           IF "CNV_HMI".Charge_Commands[#HMI_No] THEN
               CASE #"ID(1)" OF
                       //CNV 1 - SYSTEM 1
                   100101:
                       #"Enable(1)" := "Control_DB".LCnv_Sys[#Sys_No].Cnv_Level[1].Cnv1.Instruction.Enable;
                       #"Mode_Change(1)" := "Control_DB".LCnv_Sys[#Sys_No].Cnv_Level[1].Cnv1.Instruction.Mode_Change;
                       #"Transfer_To_ID(1)" := "Control_DB".LCnv_Sys[#Sys_No].Cnv_Level[1].Cnv1.Instruction.Transfer_To_ID;
                       #"Transfer_From_ID(1)" := "Control_DB".LCnv_Sys[#Sys_No].Cnv_Level[1].Cnv1.Instruction.Transfer_From_ID;
                       #"Pallet_Allignment(1)" := "Control_DB".LCnv_Sys[#Sys_No].Cnv_Level[1].Cnv1.Instruction.Pallet_Allignment;
                   100201:
                       "Enable_HMI(1)" := "Control_DB".LCnv_Sys[#Sys_No].Cnv_Level[2].Cnv1.Instruction.Enable;
                       "Mode_Change_HMI(1)" := "Control_DB".LCnv_Sys[#Sys_No].Cnv_Level[2].Cnv1.Instruction.Mode_Change;
                       "Transfer_To_ID_HMI(1)" := "Control_DB".LCnv_Sys[#Sys_No].Cnv_Level[2].Cnv1.Instruction.Transfer_To_ID;
                       "Transfer_From_ID_HMI(1)" := "Control_DB".LCnv_Sys[#Sys_No].Cnv_Level[2].Cnv1.Instruction.Transfer_From_ID;
                       "Pallet_Allignment_HMI(1)" := "Control_DB".LCnv_Sys[#Sys_No].Cnv_Level[2].Cnv1.Instruction.Pallet_Allignment;
                   100301:
                       "Enable_HMI(1)" := "Control_DB".LCnv_Sys[#Sys_No].Cnv_Level[3].Cnv1.Instruction.Enable;
                       "Mode_Change_HMI(1)" := "Control_DB".LCnv_Sys[#Sys_No].Cnv_Level[3].Cnv1.Instruction.Mode_Change;
                       "Transfer_To_ID_HMI(1)" := "Control_DB".LCnv_Sys[#Sys_No].Cnv_Level[3].Cnv1.Instruction.Transfer_To_ID;
                       "Transfer_From_ID_HMI(1)" := "Control_DB".LCnv_Sys[#Sys_No].Cnv_Level[3].Cnv1.Instruction.Transfer_From_ID;
                       "Pallet_Allignment_HMI(1)" := "Control_DB".LCnv_Sys[#Sys_No].Cnv_Level[3].Cnv1.Instruction.Pallet_Allignment;
                   100401:
                       "Enable_HMI(1)" := "Control_DB".LCnv_Sys[#Sys_No].Cnv_Level[4].Cnv1.Instruction.Enable;
                       "Mode_Change_HMI(1)" := "Control_DB".LCnv_Sys[#Sys_No].Cnv_Level[4].Cnv1.Instruction.Mode_Change;
                       "Transfer_To_ID_HMI(1)" := "Control_DB".LCnv_Sys[#Sys_No].Cnv_Level[4].Cnv1.Instruction.Transfer_To_ID;
                       "Transfer_From_ID_HMI(1)" := "Control_DB".LCnv_Sys[#Sys_No].Cnv_Level[4].Cnv1.Instruction.Transfer_From_ID;
                       "Pallet_Allignment_HMI(1)" := "Control_DB".LCnv_Sys[#Sys_No].Cnv_Level[4].Cnv1.Instruction.Pallet_Allignment;
                   100501:
                       "Enable_HMI(1)" := "Control_DB".LCnv_Sys[#Sys_No].Cnv_Level[5].Cnv1.Instruction.Enable;
                       "Mode_Change_HMI(1)" := "Control_DB".LCnv_Sys[#Sys_No].Cnv_Level[5].Cnv1.Instruction.Mode_Change;
                       "Task_ID_HMI(1)" := "Control_DB".LCnv_Sys[#Sys_No].Cnv_Level[5].Cnv1.Instruction.Task_ID;
                       "Transfer_To_ID_HMI(1)" := "Control_DB".LCnv_Sys[#Sys_No].Cnv_Level[5].Cnv1.Instruction.Transfer_To_ID;
                       "Transfer_From_ID_HMI(1)" := "Control_DB".LCnv_Sys[#Sys_No].Cnv_Level[5].Cnv1.Instruction.Transfer_From_ID;
                       "Pallet_Allignment_HMI(1)" := "Control_DB".LCnv_Sys[#Sys_No].Cnv_Level[5].Cnv1.Instruction.Pallet_Allignment;
                   100601:
                       "Enable_HMI(1)" := "Control_DB".LCnv_Sys[#Sys_No].Cnv_Level[6].Cnv1.Instruction.Enable;
                       "Mode_Change_HMI(1)" := "Control_DB".LCnv_Sys[#Sys_No].Cnv_Level[6].Cnv1.Instruction.Mode_Change;
                       "Task_ID_HMI(1)" := "Control_DB".LCnv_Sys[#Sys_No].Cnv_Level[6].Cnv1.Instruction.Task_ID;
                       "Transfer_To_ID_HMI(1)" := "Control_DB".LCnv_Sys[#Sys_No].Cnv_Level[6].Cnv1.Instruction.Transfer_To_ID;
                       "Transfer_From_ID_HMI(1)" := "Control_DB".LCnv_Sys[#Sys_No].Cnv_Level[6].Cnv1.Instruction.Transfer_From_ID;
                       "Pallet_Allignment_HMI(1)" := "Control_DB".LCnv_Sys[#Sys_No].Cnv_Level[6].Cnv1.Instruction.Pallet_Allignment;
                   100701:
                       "Enable_HMI(1)" := "Control_DB".LCnv_Sys[#Sys_No].Cnv_Level[7].Cnv1.Instruction.Enable;
                       "Mode_Change_HMI(1)" := "Control_DB".LCnv_Sys[#Sys_No].Cnv_Level[7].Cnv1.Instruction.Mode_Change;
                       "Task_ID_HMI(1)" := "Control_DB".LCnv_Sys[#Sys_No].Cnv_Level[7].Cnv1.Instruction.Task_ID;
                       "Transfer_To_ID_HMI(1)" := "Control_DB".LCnv_Sys[#Sys_No].Cnv_Level[7].Cnv1.Instruction.Transfer_To_ID;
                       "Transfer_From_ID_HMI(1)" := "Control_DB".LCnv_Sys[#Sys_No].Cnv_Level[7].Cnv1.Instruction.Transfer_From_ID;
                       "Pallet_Allignment_HMI(1)" := "Control_DB".LCnv_Sys[#Sys_No].Cnv_Level[7].Cnv1.Instruction.Pallet_Allignment;
                   100801:
                       "Enable_HMI(1)" := "Control_DB".LCnv_Sys[#Sys_No].Cnv_Level[8].Cnv1.Instruction.Enable;
                       "Mode_Change_HMI(1)" := "Control_DB".LCnv_Sys[#Sys_No].Cnv_Level[8].Cnv1.Instruction.Mode_Change;
                       "Task_ID_HMI(1)" := "Control_DB".LCnv_Sys[#Sys_No].Cnv_Level[8].Cnv1.Instruction.Task_ID;
                       "Transfer_To_ID_HMI(1)" := "Control_DB".LCnv_Sys[#Sys_No].Cnv_Level[8].Cnv1.Instruction.Transfer_To_ID;
                       "Transfer_From_ID_HMI(1)" := "Control_DB".LCnv_Sys[#Sys_No].Cnv_Level[8].Cnv1.Instruction.Transfer_From_ID;
                       "Pallet_Allignment_HMI(1)" := "Control_DB".LCnv_Sys[#Sys_No].Cnv_Level[8].Cnv1.Instruction.Pallet_Allignment;
                       //CNV 2 - SYSTEM 1
                   110101:
                       "Enable_HMI(1)" := "Control_DB".LCnv_Sys[#Sys_No].Cnv_Level[1].Cnv2.Instruction.Enable;
                       "Mode_Change_HMI(1)" := "Control_DB".LCnv_Sys[#Sys_No].Cnv_Level[1].Cnv2.Instruction.Mode_Change;
                       "Task_ID_HMI(1)" := "Control_DB".LCnv_Sys[#Sys_No].Cnv_Level[1].Cnv2.Instruction.Task_ID;
                       "Transfer_To_ID_HMI(1)" := "Control_DB".LCnv_Sys[#Sys_No].Cnv_Level[1].Cnv2.Instruction.Transfer_To_ID;
                       "Transfer_From_ID_HMI(1)" := "Control_DB".LCnv_Sys[#Sys_No].Cnv_Level[1].Cnv2.Instruction.Transfer_From_ID;
                       "Pallet_Allignment_HMI(1)" := "Control_DB".LCnv_Sys[#Sys_No].Cnv_Level[1].Cnv2.Instruction.Pallet_Allignment;
                   110201:
                       "Enable_HMI(1)" := "Control_DB".LCnv_Sys[#Sys_No].Cnv_Level[2].Cnv2.Instruction.Enable;
                       "Mode_Change_HMI(1)" := "Control_DB".LCnv_Sys[#Sys_No].Cnv_Level[2].Cnv2.Instruction.Mode_Change;
                       "Task_ID_HMI(1)" := "Control_DB".LCnv_Sys[#Sys_No].Cnv_Level[2].Cnv2.Instruction.Task_ID;
                       "Transfer_To_ID_HMI(1)" := "Control_DB".LCnv_Sys[#Sys_No].Cnv_Level[2].Cnv2.Instruction.Transfer_To_ID;
                       "Transfer_From_ID_HMI(1)" := "Control_DB".LCnv_Sys[#Sys_No].Cnv_Level[2].Cnv2.Instruction.Transfer_From_ID;
                       "Pallet_Allignment_HMI(1)" := "Control_DB".LCnv_Sys[#Sys_No].Cnv_Level[2].Cnv2.Instruction.Pallet_Allignment;
                   110301:
                       "Enable_HMI(1)" := "Control_DB".LCnv_Sys[#Sys_No].Cnv_Level[3].Cnv2.Instruction.Enable;
                       "Mode_Change_HMI(1)" := "Control_DB".LCnv_Sys[#Sys_No].Cnv_Level[3].Cnv2.Instruction.Mode_Change;
                       "Task_ID_HMI(1)" := "Control_DB".LCnv_Sys[#Sys_No].Cnv_Level[3].Cnv2.Instruction.Task_ID;
                       "Transfer_To_ID_HMI(1)" := "Control_DB".LCnv_Sys[#Sys_No].Cnv_Level[3].Cnv2.Instruction.Transfer_To_ID;
                       "Transfer_From_ID_HMI(1)" := "Control_DB".LCnv_Sys[#Sys_No].Cnv_Level[3].Cnv2.Instruction.Transfer_From_ID;
                       "Pallet_Allignment_HMI(1)" := "Control_DB".LCnv_Sys[#Sys_No].Cnv_Level[3].Cnv2.Instruction.Pallet_Allignment;
                   110401:
                       "Enable_HMI(1)" := "Control_DB".LCnv_Sys[#Sys_No].Cnv_Level[4].Cnv2.Instruction.Enable;
                       "Mode_Change_HMI(1)" := "Control_DB".LCnv_Sys[#Sys_No].Cnv_Level[4].Cnv2.Instruction.Mode_Change;
                       "Task_ID_HMI(1)" := "Control_DB".LCnv_Sys[#Sys_No].Cnv_Level[4].Cnv2.Instruction.Task_ID;
                       "Transfer_To_ID_HMI(1)" := "Control_DB".LCnv_Sys[#Sys_No].Cnv_Level[4].Cnv2.Instruction.Transfer_To_ID;
                       "Transfer_From_ID_HMI(1)" := "Control_DB".LCnv_Sys[#Sys_No].Cnv_Level[4].Cnv2.Instruction.Transfer_From_ID;
                       "Pallet_Allignment_HMI(1)" := "Control_DB".LCnv_Sys[#Sys_No].Cnv_Level[4].Cnv2.Instruction.Pallet_Allignment;
                   110501:
                       "Enable_HMI(1)" := "Control_DB".LCnv_Sys[#Sys_No].Cnv_Level[5].Cnv2.Instruction.Enable;
                       "Mode_Change_HMI(1)" := "Control_DB".LCnv_Sys[#Sys_No].Cnv_Level[5].Cnv2.Instruction.Mode_Change;
                       "Task_ID_HMI(1)" := "Control_DB".LCnv_Sys[#Sys_No].Cnv_Level[5].Cnv2.Instruction.Task_ID;
                       "Transfer_To_ID_HMI(1)" := "Control_DB".LCnv_Sys[#Sys_No].Cnv_Level[5].Cnv2.Instruction.Transfer_To_ID;
                       "Transfer_From_ID_HMI(1)" := "Control_DB".LCnv_Sys[#Sys_No].Cnv_Level[5].Cnv2.Instruction.Transfer_From_ID;
                       "Pallet_Allignment_HMI(1)" := "Control_DB".LCnv_Sys[#Sys_No].Cnv_Level[5].Cnv2.Instruction.Pallet_Allignment;
                   110601:
                       "Enable_HMI(1)" := "Control_DB".LCnv_Sys[#Sys_No].Cnv_Level[6].Cnv2.Instruction.Enable;
                       "Mode_Change_HMI(1)" := "Control_DB".LCnv_Sys[#Sys_No].Cnv_Level[6].Cnv2.Instruction.Mode_Change;
                       "Task_ID_HMI(1)" := "Control_DB".LCnv_Sys[#Sys_No].Cnv_Level[6].Cnv2.Instruction.Task_ID;
                       "Transfer_To_ID_HMI(1)" := "Control_DB".LCnv_Sys[#Sys_No].Cnv_Level[6].Cnv2.Instruction.Transfer_To_ID;
                       "Transfer_From_ID_HMI(1)" := "Control_DB".LCnv_Sys[#Sys_No].Cnv_Level[6].Cnv2.Instruction.Transfer_From_ID;
                       "Pallet_Allignment_HMI(1)" := "Control_DB".LCnv_Sys[#Sys_No].Cnv_Level[6].Cnv2.Instruction.Pallet_Allignment;
                   110701:
                       "Enable_HMI(1)" := "Control_DB".LCnv_Sys[#Sys_No].Cnv_Level[7].Cnv2.Instruction.Enable;
                       "Mode_Change_HMI(1)" := "Control_DB".LCnv_Sys[#Sys_No].Cnv_Level[7].Cnv2.Instruction.Mode_Change;
                       "Task_ID_HMI(1)" := "Control_DB".LCnv_Sys[#Sys_No].Cnv_Level[7].Cnv2.Instruction.Task_ID;
                       "Transfer_To_ID_HMI(1)" := "Control_DB".LCnv_Sys[#Sys_No].Cnv_Level[7].Cnv2.Instruction.Transfer_To_ID;
                       "Transfer_From_ID_HMI(1)" := "Control_DB".LCnv_Sys[#Sys_No].Cnv_Level[7].Cnv2.Instruction.Transfer_From_ID;
                       "Pallet_Allignment_HMI(1)" := "Control_DB".LCnv_Sys[#Sys_No].Cnv_Level[7].Cnv2.Instruction.Pallet_Allignment;
                   110801:
                       "Enable_HMI(1)" := "Control_DB".LCnv_Sys[#Sys_No].Cnv_Level[8].Cnv2.Instruction.Enable;
                       "Mode_Change_HMI(1)" := "Control_DB".LCnv_Sys[#Sys_No].Cnv_Level[8].Cnv2.Instruction.Mode_Change;
                       "Task_ID_HMI(1)" := "Control_DB".LCnv_Sys[#Sys_No].Cnv_Level[8].Cnv2.Instruction.Task_ID;
                       "Transfer_To_ID_HMI(1)" := "Control_DB".LCnv_Sys[#Sys_No].Cnv_Level[8].Cnv2.Instruction.Transfer_To_ID;
                       "Transfer_From_ID_HMI(1)" := "Control_DB".LCnv_Sys[#Sys_No].Cnv_Level[8].Cnv2.Instruction.Transfer_From_ID;
                       "Pallet_Allignment_HMI(1)" := "Control_DB".LCnv_Sys[#Sys_No].Cnv_Level[8].Cnv2.Instruction.Pallet_Allignment;
                       //CNV 1 - SYSTEM 2
                   100102:
                       "Enable_HMI(1)" := "Control_DB".LCnv_Sys[2].Cnv_Level[1].Cnv1.Instruction.Enable;
                       "Mode_Change_HMI(1)" := "Control_DB".LCnv_Sys[2].Cnv_Level[1].Cnv1.Instruction.Mode_Change;
                       "Task_ID_HMI(1)" := "Control_DB".LCnv_Sys[2].Cnv_Level[1].Cnv1.Instruction.Task_ID;
                       "Transfer_To_ID_HMI(1)" := "Control_DB".LCnv_Sys[2].Cnv_Level[1].Cnv1.Instruction.Transfer_To_ID;
                       "Transfer_From_ID_HMI(1)" := "Control_DB".LCnv_Sys[2].Cnv_Level[1].Cnv1.Instruction.Transfer_From_ID;
                       "Pallet_Allignment_HMI(1)" := "Control_DB".LCnv_Sys[2].Cnv_Level[1].Cnv1.Instruction.Pallet_Allignment;
                   100202:
                       "Enable_HMI(1)" := "Control_DB".LCnv_Sys[2].Cnv_Level[2].Cnv1.Instruction.Enable;
                       "Mode_Change_HMI(1)" := "Control_DB".LCnv_Sys[2].Cnv_Level[2].Cnv1.Instruction.Mode_Change;
                       "Task_ID_HMI(1)" := "Control_DB".LCnv_Sys[2].Cnv_Level[2].Cnv1.Instruction.Task_ID;
                       "Transfer_To_ID_HMI(1)" := "Control_DB".LCnv_Sys[2].Cnv_Level[2].Cnv1.Instruction.Transfer_To_ID;
                       "Transfer_From_ID_HMI(1)" := "Control_DB".LCnv_Sys[2].Cnv_Level[2].Cnv1.Instruction.Transfer_From_ID;
                       "Pallet_Allignment_HMI(1)" := "Control_DB".LCnv_Sys[2].Cnv_Level[2].Cnv1.Instruction.Pallet_Allignment;
                   100302:
                       "Enable_HMI(1)" := "Control_DB".LCnv_Sys[2].Cnv_Level[3].Cnv1.Instruction.Enable;
                       "Mode_Change_HMI(1)" := "Control_DB".LCnv_Sys[2].Cnv_Level[3].Cnv1.Instruction.Mode_Change;
                       "Task_ID_HMI(1)" := "Control_DB".LCnv_Sys[2].Cnv_Level[3].Cnv1.Instruction.Task_ID;
                       "Transfer_To_ID_HMI(1)" := "Control_DB".LCnv_Sys[2].Cnv_Level[3].Cnv1.Instruction.Transfer_To_ID;
                       "Transfer_From_ID_HMI(1)" := "Control_DB".LCnv_Sys[2].Cnv_Level[3].Cnv1.Instruction.Transfer_From_ID;
                       "Pallet_Allignment_HMI(1)" := "Control_DB".LCnv_Sys[2].Cnv_Level[3].Cnv1.Instruction.Pallet_Allignment;
                   100402:
                       "Enable_HMI(1)" := "Control_DB".LCnv_Sys[2].Cnv_Level[4].Cnv1.Instruction.Enable;
                       "Mode_Change_HMI(1)" := "Control_DB".LCnv_Sys[2].Cnv_Level[4].Cnv1.Instruction.Mode_Change;
                       "Task_ID_HMI(1)" := "Control_DB".LCnv_Sys[2].Cnv_Level[4].Cnv1.Instruction.Task_ID;
                       "Transfer_To_ID_HMI(1)" := "Control_DB".LCnv_Sys[2].Cnv_Level[4].Cnv1.Instruction.Transfer_To_ID;
                       "Transfer_From_ID_HMI(1)" := "Control_DB".LCnv_Sys[2].Cnv_Level[4].Cnv1.Instruction.Transfer_From_ID;
                       "Pallet_Allignment_HMI(1)" := "Control_DB".LCnv_Sys[2].Cnv_Level[4].Cnv1.Instruction.Pallet_Allignment;
                   100502:
                       "Enable_HMI(1)" := "Control_DB".LCnv_Sys[2].Cnv_Level[5].Cnv1.Instruction.Enable;
                       "Mode_Change_HMI(1)" := "Control_DB".LCnv_Sys[2].Cnv_Level[5].Cnv1.Instruction.Mode_Change;
                       "Task_ID_HMI(1)" := "Control_DB".LCnv_Sys[2].Cnv_Level[5].Cnv1.Instruction.Task_ID;
                       "Transfer_To_ID_HMI(1)" := "Control_DB".LCnv_Sys[2].Cnv_Level[5].Cnv1.Instruction.Transfer_To_ID;
                       "Transfer_From_ID_HMI(1)" := "Control_DB".LCnv_Sys[2].Cnv_Level[5].Cnv1.Instruction.Transfer_From_ID;
                       "Pallet_Allignment_HMI(1)" := "Control_DB".LCnv_Sys[2].Cnv_Level[5].Cnv1.Instruction.Pallet_Allignment;
                   100602:
                       "Enable_HMI(1)" := "Control_DB".LCnv_Sys[2].Cnv_Level[6].Cnv1.Instruction.Enable;
                       "Mode_Change_HMI(1)" := "Control_DB".LCnv_Sys[2].Cnv_Level[6].Cnv1.Instruction.Mode_Change;
                       "Task_ID_HMI(1)" := "Control_DB".LCnv_Sys[2].Cnv_Level[6].Cnv1.Instruction.Task_ID;
                       "Transfer_To_ID_HMI(1)" := "Control_DB".LCnv_Sys[2].Cnv_Level[6].Cnv1.Instruction.Transfer_To_ID;
                       "Transfer_From_ID_HMI(1)" := "Control_DB".LCnv_Sys[2].Cnv_Level[6].Cnv1.Instruction.Transfer_From_ID;
                       "Pallet_Allignment_HMI(1)" := "Control_DB".LCnv_Sys[2].Cnv_Level[6].Cnv1.Instruction.Pallet_Allignment;
                   100702:
                       "Enable_HMI(1)" := "Control_DB".LCnv_Sys[2].Cnv_Level[7].Cnv1.Instruction.Enable;
                       "Mode_Change_HMI(1)" := "Control_DB".LCnv_Sys[2].Cnv_Level[7].Cnv1.Instruction.Mode_Change;
                       "Task_ID_HMI(1)" := "Control_DB".LCnv_Sys[2].Cnv_Level[7].Cnv1.Instruction.Task_ID;
                       "Transfer_To_ID_HMI(1)" := "Control_DB".LCnv_Sys[2].Cnv_Level[7].Cnv1.Instruction.Transfer_To_ID;
                       "Transfer_From_ID_HMI(1)" := "Control_DB".LCnv_Sys[2].Cnv_Level[7].Cnv1.Instruction.Transfer_From_ID;
                       "Pallet_Allignment_HMI(1)" := "Control_DB".LCnv_Sys[2].Cnv_Level[7].Cnv1.Instruction.Pallet_Allignment;
                   100802:
                       "Enable_HMI(1)" := "Control_DB".LCnv_Sys[2].Cnv_Level[8].Cnv1.Instruction.Enable;
                       "Mode_Change_HMI(1)" := "Control_DB".LCnv_Sys[2].Cnv_Level[8].Cnv1.Instruction.Mode_Change;
                       "Task_ID_HMI(1)" := "Control_DB".LCnv_Sys[2].Cnv_Level[8].Cnv1.Instruction.Task_ID;
                       "Transfer_To_ID_HMI(1)" := "Control_DB".LCnv_Sys[2].Cnv_Level[8].Cnv1.Instruction.Transfer_To_ID;
                       "Transfer_From_ID_HMI(1)" := "Control_DB".LCnv_Sys[2].Cnv_Level[8].Cnv1.Instruction.Transfer_From_ID;
                       "Pallet_Allignment_HMI(1)" := "Control_DB".LCnv_Sys[2].Cnv_Level[8].Cnv1.Instruction.Pallet_Allignment;
                       //CNV 2 - SYSTEM 2
                   110102:
                       "Enable_HMI(1)" := "Control_DB".LCnv_Sys[2].Cnv_Level[1].Cnv2.Instruction.Enable;
                       "Mode_Change_HMI(1)" := "Control_DB".LCnv_Sys[2].Cnv_Level[1].Cnv2.Instruction.Mode_Change;
                       "Task_ID_HMI(1)" := "Control_DB".LCnv_Sys[2].Cnv_Level[1].Cnv2.Instruction.Task_ID;
                       "Transfer_To_ID_HMI(1)" := "Control_DB".LCnv_Sys[2].Cnv_Level[1].Cnv2.Instruction.Transfer_To_ID;
                       "Transfer_From_ID_HMI(1)" := "Control_DB".LCnv_Sys[2].Cnv_Level[1].Cnv2.Instruction.Transfer_From_ID;
                       "Pallet_Allignment_HMI(1)" := "Control_DB".LCnv_Sys[2].Cnv_Level[1].Cnv2.Instruction.Pallet_Allignment;
                   110202:
                       "Enable_HMI(1)" := "Control_DB".LCnv_Sys[2].Cnv_Level[2].Cnv2.Instruction.Enable;
                       "Mode_Change_HMI(1)" := "Control_DB".LCnv_Sys[2].Cnv_Level[2].Cnv2.Instruction.Mode_Change;
                       "Task_ID_HMI(1)" := "Control_DB".LCnv_Sys[2].Cnv_Level[2].Cnv2.Instruction.Task_ID;
                       "Transfer_To_ID_HMI(1)" := "Control_DB".LCnv_Sys[2].Cnv_Level[2].Cnv2.Instruction.Transfer_To_ID;
                       "Transfer_From_ID_HMI(1)" := "Control_DB".LCnv_Sys[2].Cnv_Level[2].Cnv2.Instruction.Transfer_From_ID;
                       "Pallet_Allignment_HMI(1)" := "Control_DB".LCnv_Sys[2].Cnv_Level[2].Cnv2.Instruction.Pallet_Allignment;
                   110302:
                       "Enable_HMI(1)" := "Control_DB".LCnv_Sys[2].Cnv_Level[3].Cnv2.Instruction.Enable;
                       "Mode_Change_HMI(1)" := "Control_DB".LCnv_Sys[2].Cnv_Level[3].Cnv2.Instruction.Mode_Change;
                       "Task_ID_HMI(1)" := "Control_DB".LCnv_Sys[2].Cnv_Level[3].Cnv2.Instruction.Task_ID;
                       "Transfer_To_ID_HMI(1)" := "Control_DB".LCnv_Sys[2].Cnv_Level[3].Cnv2.Instruction.Transfer_To_ID;
                       "Transfer_From_ID_HMI(1)" := "Control_DB".LCnv_Sys[2].Cnv_Level[3].Cnv2.Instruction.Transfer_From_ID;
                       "Pallet_Allignment_HMI(1)" := "Control_DB".LCnv_Sys[2].Cnv_Level[3].Cnv2.Instruction.Pallet_Allignment;
                   110402:
                       "Enable_HMI(1)" := "Control_DB".LCnv_Sys[2].Cnv_Level[4].Cnv2.Instruction.Enable;
                       "Mode_Change_HMI(1)" := "Control_DB".LCnv_Sys[2].Cnv_Level[4].Cnv2.Instruction.Mode_Change;
                       "Task_ID_HMI(1)" := "Control_DB".LCnv_Sys[2].Cnv_Level[4].Cnv2.Instruction.Task_ID;
                       "Transfer_To_ID_HMI(1)" := "Control_DB".LCnv_Sys[2].Cnv_Level[4].Cnv2.Instruction.Transfer_To_ID;
                       "Transfer_From_ID_HMI(1)" := "Control_DB".LCnv_Sys[2].Cnv_Level[4].Cnv2.Instruction.Transfer_From_ID;
                       "Pallet_Allignment_HMI(1)" := "Control_DB".LCnv_Sys[2].Cnv_Level[4].Cnv2.Instruction.Pallet_Allignment;
                   110502:
                       "Enable_HMI(1)" := "Control_DB".LCnv_Sys[2].Cnv_Level[5].Cnv2.Instruction.Enable;
                       "Mode_Change_HMI(1)" := "Control_DB".LCnv_Sys[2].Cnv_Level[5].Cnv2.Instruction.Mode_Change;
                       "Task_ID_HMI(1)" := "Control_DB".LCnv_Sys[2].Cnv_Level[5].Cnv2.Instruction.Task_ID;
                       "Transfer_To_ID_HMI(1)" := "Control_DB".LCnv_Sys[2].Cnv_Level[5].Cnv2.Instruction.Transfer_To_ID;
                       "Transfer_From_ID_HMI(1)" := "Control_DB".LCnv_Sys[2].Cnv_Level[5].Cnv2.Instruction.Transfer_From_ID;
                       "Pallet_Allignment_HMI(1)" := "Control_DB".LCnv_Sys[2].Cnv_Level[5].Cnv2.Instruction.Pallet_Allignment;
                   110602:
                       "Enable_HMI(1)" := "Control_DB".LCnv_Sys[2].Cnv_Level[6].Cnv2.Instruction.Enable;
                       "Mode_Change_HMI(1)" := "Control_DB".LCnv_Sys[2].Cnv_Level[6].Cnv2.Instruction.Mode_Change;
                       "Task_ID_HMI(1)" := "Control_DB".LCnv_Sys[2].Cnv_Level[6].Cnv2.Instruction.Task_ID;
                       "Transfer_To_ID_HMI(1)" := "Control_DB".LCnv_Sys[2].Cnv_Level[6].Cnv2.Instruction.Transfer_To_ID;
                       "Transfer_From_ID_HMI(1)" := "Control_DB".LCnv_Sys[2].Cnv_Level[6].Cnv2.Instruction.Transfer_From_ID;
                       "Pallet_Allignment_HMI(1)" := "Control_DB".LCnv_Sys[2].Cnv_Level[6].Cnv2.Instruction.Pallet_Allignment;
                   110702:
                       "Enable_HMI(1)" := "Control_DB".LCnv_Sys[2].Cnv_Level[7].Cnv2.Instruction.Enable;
                       "Mode_Change_HMI(1)" := "Control_DB".LCnv_Sys[2].Cnv_Level[7].Cnv2.Instruction.Mode_Change;
                       "Task_ID_HMI(1)" := "Control_DB".LCnv_Sys[2].Cnv_Level[7].Cnv2.Instruction.Task_ID;
                       "Transfer_To_ID_HMI(1)" := "Control_DB".LCnv_Sys[2].Cnv_Level[7].Cnv2.Instruction.Transfer_To_ID;
                       "Transfer_From_ID_HMI(1)" := "Control_DB".LCnv_Sys[2].Cnv_Level[7].Cnv2.Instruction.Transfer_From_ID;
                       "Pallet_Allignment_HMI(1)" := "Control_DB".LCnv_Sys[2].Cnv_Level[7].Cnv2.Instruction.Pallet_Allignment;
                   110802:
                       "Enable_HMI(1)" := "Control_DB".LCnv_Sys[2].Cnv_Level[8].Cnv2.Instruction.Enable;
                       "Mode_Change_HMI(1)" := "Control_DB".LCnv_Sys[2].Cnv_Level[8].Cnv2.Instruction.Mode_Change;
                       "Task_ID_HMI(1)" := "Control_DB".LCnv_Sys[2].Cnv_Level[8].Cnv2.Instruction.Task_ID;
                       "Transfer_To_ID_HMI(1)" := "Control_DB".LCnv_Sys[2].Cnv_Level[8].Cnv2.Instruction.Transfer_To_ID;
                       "Transfer_From_ID_HMI(1)" := "Control_DB".LCnv_Sys[2].Cnv_Level[8].Cnv2.Instruction.Transfer_From_ID;
                       "Pallet_Allignment_HMI(1)" := "Control_DB".LCnv_Sys[2].Cnv_Level[8].Cnv2.Instruction.Pallet_Allignment;
                       //CNV 1 - SYSTEM 3
                   100103:
                       "Enable_HMI(1)" := "Control_DB".LCnv_Sys[3].Cnv_Level[1].Cnv1.Instruction.Enable;
                       "Mode_Change_HMI(1)" := "Control_DB".LCnv_Sys[3].Cnv_Level[1].Cnv1.Instruction.Mode_Change;
                       "Task_ID_HMI(1)" := "Control_DB".LCnv_Sys[3].Cnv_Level[1].Cnv1.Instruction.Task_ID;
                       "Transfer_To_ID_HMI(1)" := "Control_DB".LCnv_Sys[3].Cnv_Level[1].Cnv1.Instruction.Transfer_To_ID;
                       "Transfer_From_ID_HMI(1)" := "Control_DB".LCnv_Sys[3].Cnv_Level[1].Cnv1.Instruction.Transfer_From_ID;
                       "Pallet_Allignment_HMI(1)" := "Control_DB".LCnv_Sys[3].Cnv_Level[1].Cnv1.Instruction.Pallet_Allignment;
                   100203:
                       "Enable_HMI(1)" := "Control_DB".LCnv_Sys[3].Cnv_Level[2].Cnv1.Instruction.Enable;
                       "Mode_Change_HMI(1)" := "Control_DB".LCnv_Sys[3].Cnv_Level[2].Cnv1.Instruction.Mode_Change;
                       "Task_ID_HMI(1)" := "Control_DB".LCnv_Sys[3].Cnv_Level[2].Cnv1.Instruction.Task_ID;
                       "Transfer_To_ID_HMI(1)" := "Control_DB".LCnv_Sys[3].Cnv_Level[2].Cnv1.Instruction.Transfer_To_ID;
                       "Transfer_From_ID_HMI(1)" := "Control_DB".LCnv_Sys[3].Cnv_Level[2].Cnv1.Instruction.Transfer_From_ID;
                       "Pallet_Allignment_HMI(1)" := "Control_DB".LCnv_Sys[3].Cnv_Level[2].Cnv1.Instruction.Pallet_Allignment;
                   100303:
                       "Enable_HMI(1)" := "Control_DB".LCnv_Sys[3].Cnv_Level[3].Cnv1.Instruction.Enable;
                       "Mode_Change_HMI(1)" := "Control_DB".LCnv_Sys[3].Cnv_Level[3].Cnv1.Instruction.Mode_Change;
                       "Task_ID_HMI(1)" := "Control_DB".LCnv_Sys[3].Cnv_Level[3].Cnv1.Instruction.Task_ID;
                       "Transfer_To_ID_HMI(1)" := "Control_DB".LCnv_Sys[3].Cnv_Level[3].Cnv1.Instruction.Transfer_To_ID;
                       "Transfer_From_ID_HMI(1)" := "Control_DB".LCnv_Sys[3].Cnv_Level[3].Cnv1.Instruction.Transfer_From_ID;
                       "Pallet_Allignment_HMI(1)" := "Control_DB".LCnv_Sys[3].Cnv_Level[3].Cnv1.Instruction.Pallet_Allignment;
                   100403:
                       "Enable_HMI(1)" := "Control_DB".LCnv_Sys[3].Cnv_Level[4].Cnv1.Instruction.Enable;
                       "Mode_Change_HMI(1)" := "Control_DB".LCnv_Sys[3].Cnv_Level[4].Cnv1.Instruction.Mode_Change;
                       "Task_ID_HMI(1)" := "Control_DB".LCnv_Sys[3].Cnv_Level[4].Cnv1.Instruction.Task_ID;
                       "Transfer_To_ID_HMI(1)" := "Control_DB".LCnv_Sys[3].Cnv_Level[4].Cnv1.Instruction.Transfer_To_ID;
                       "Transfer_From_ID_HMI(1)" := "Control_DB".LCnv_Sys[3].Cnv_Level[4].Cnv1.Instruction.Transfer_From_ID;
                       "Pallet_Allignment_HMI(1)" := "Control_DB".LCnv_Sys[3].Cnv_Level[4].Cnv1.Instruction.Pallet_Allignment;
                   100503:
                       "Enable_HMI(1)" := "Control_DB".LCnv_Sys[3].Cnv_Level[5].Cnv1.Instruction.Enable;
                       "Mode_Change_HMI(1)" := "Control_DB".LCnv_Sys[3].Cnv_Level[5].Cnv1.Instruction.Mode_Change;
                       "Task_ID_HMI(1)" := "Control_DB".LCnv_Sys[3].Cnv_Level[5].Cnv1.Instruction.Task_ID;
                       "Transfer_To_ID_HMI(1)" := "Control_DB".LCnv_Sys[3].Cnv_Level[5].Cnv1.Instruction.Transfer_To_ID;
                       "Transfer_From_ID_HMI(1)" := "Control_DB".LCnv_Sys[3].Cnv_Level[5].Cnv1.Instruction.Transfer_From_ID;
                       "Pallet_Allignment_HMI(1)" := "Control_DB".LCnv_Sys[3].Cnv_Level[5].Cnv1.Instruction.Pallet_Allignment;
                   100603:
                       "Enable_HMI(1)" := "Control_DB".LCnv_Sys[3].Cnv_Level[6].Cnv1.Instruction.Enable;
                       "Mode_Change_HMI(1)" := "Control_DB".LCnv_Sys[3].Cnv_Level[6].Cnv1.Instruction.Mode_Change;
                       "Task_ID_HMI(1)" := "Control_DB".LCnv_Sys[3].Cnv_Level[6].Cnv1.Instruction.Task_ID;
                       "Transfer_To_ID_HMI(1)" := "Control_DB".LCnv_Sys[3].Cnv_Level[6].Cnv1.Instruction.Transfer_To_ID;
                       "Transfer_From_ID_HMI(1)" := "Control_DB".LCnv_Sys[3].Cnv_Level[6].Cnv1.Instruction.Transfer_From_ID;
                       "Pallet_Allignment_HMI(1)" := "Control_DB".LCnv_Sys[3].Cnv_Level[6].Cnv1.Instruction.Pallet_Allignment;
                   100703:
                       "Enable_HMI(1)" := "Control_DB".LCnv_Sys[3].Cnv_Level[7].Cnv1.Instruction.Enable;
                       "Mode_Change_HMI(1)" := "Control_DB".LCnv_Sys[3].Cnv_Level[7].Cnv1.Instruction.Mode_Change;
                       "Task_ID_HMI(1)" := "Control_DB".LCnv_Sys[3].Cnv_Level[7].Cnv1.Instruction.Task_ID;
                       "Transfer_To_ID_HMI(1)" := "Control_DB".LCnv_Sys[3].Cnv_Level[7].Cnv1.Instruction.Transfer_To_ID;
                       "Transfer_From_ID_HMI(1)" := "Control_DB".LCnv_Sys[3].Cnv_Level[7].Cnv1.Instruction.Transfer_From_ID;
                       "Pallet_Allignment_HMI(1)" := "Control_DB".LCnv_Sys[3].Cnv_Level[7].Cnv1.Instruction.Pallet_Allignment;
                   100803:
                       "Enable_HMI(1)" := "Control_DB".LCnv_Sys[3].Cnv_Level[8].Cnv1.Instruction.Enable;
                       "Mode_Change_HMI(1)" := "Control_DB".LCnv_Sys[3].Cnv_Level[8].Cnv1.Instruction.Mode_Change;
                       "Task_ID_HMI(1)" := "Control_DB".LCnv_Sys[3].Cnv_Level[8].Cnv1.Instruction.Task_ID;
                       "Transfer_To_ID_HMI(1)" := "Control_DB".LCnv_Sys[3].Cnv_Level[8].Cnv1.Instruction.Transfer_To_ID;
                       "Transfer_From_ID_HMI(1)" := "Control_DB".LCnv_Sys[3].Cnv_Level[8].Cnv1.Instruction.Transfer_From_ID;
                       "Pallet_Allignment_HMI(1)" := "Control_DB".LCnv_Sys[3].Cnv_Level[8].Cnv1.Instruction.Pallet_Allignment;
                       //CNV 2 - SYSTEM 3
                   110103:
                       "Enable_HMI(1)" := "Control_DB".LCnv_Sys[3].Cnv_Level[1].Cnv2.Instruction.Enable;
                       "Mode_Change_HMI(1)" := "Control_DB".LCnv_Sys[3].Cnv_Level[1].Cnv2.Instruction.Mode_Change;
                       "Task_ID_HMI(1)" := "Control_DB".LCnv_Sys[3].Cnv_Level[1].Cnv2.Instruction.Task_ID;
                       "Transfer_To_ID_HMI(1)" := "Control_DB".LCnv_Sys[3].Cnv_Level[1].Cnv2.Instruction.Transfer_To_ID;
                       "Transfer_From_ID_HMI(1)" := "Control_DB".LCnv_Sys[3].Cnv_Level[1].Cnv2.Instruction.Transfer_From_ID;
                       "Pallet_Allignment_HMI(1)" := "Control_DB".LCnv_Sys[3].Cnv_Level[1].Cnv2.Instruction.Pallet_Allignment;
                   110203:
                       "Enable_HMI(1)" := "Control_DB".LCnv_Sys[3].Cnv_Level[2].Cnv2.Instruction.Enable;
                       "Mode_Change_HMI(1)" := "Control_DB".LCnv_Sys[3].Cnv_Level[2].Cnv2.Instruction.Mode_Change;
                       "Task_ID_HMI(1)" := "Control_DB".LCnv_Sys[3].Cnv_Level[2].Cnv2.Instruction.Task_ID;
                       "Transfer_To_ID_HMI(1)" := "Control_DB".LCnv_Sys[3].Cnv_Level[2].Cnv2.Instruction.Transfer_To_ID;
                       "Transfer_From_ID_HMI(1)" := "Control_DB".LCnv_Sys[3].Cnv_Level[2].Cnv2.Instruction.Transfer_From_ID;
                       "Pallet_Allignment_HMI(1)" := "Control_DB".LCnv_Sys[3].Cnv_Level[2].Cnv2.Instruction.Pallet_Allignment;
                   110303:
                       "Enable_HMI(1)" := "Control_DB".LCnv_Sys[3].Cnv_Level[3].Cnv2.Instruction.Enable;
                       "Mode_Change_HMI(1)" := "Control_DB".LCnv_Sys[3].Cnv_Level[3].Cnv2.Instruction.Mode_Change;
                       "Task_ID_HMI(1)" := "Control_DB".LCnv_Sys[3].Cnv_Level[3].Cnv2.Instruction.Task_ID;
                       "Transfer_To_ID_HMI(1)" := "Control_DB".LCnv_Sys[3].Cnv_Level[3].Cnv2.Instruction.Transfer_To_ID;
                       "Transfer_From_ID_HMI(1)" := "Control_DB".LCnv_Sys[3].Cnv_Level[3].Cnv2.Instruction.Transfer_From_ID;
                       "Pallet_Allignment_HMI(1)" := "Control_DB".LCnv_Sys[3].Cnv_Level[3].Cnv2.Instruction.Pallet_Allignment;
                   110403:
                       "Enable_HMI(1)" := "Control_DB".LCnv_Sys[3].Cnv_Level[4].Cnv2.Instruction.Enable;
                       "Mode_Change_HMI(1)" := "Control_DB".LCnv_Sys[3].Cnv_Level[4].Cnv2.Instruction.Mode_Change;
                       "Task_ID_HMI(1)" := "Control_DB".LCnv_Sys[3].Cnv_Level[4].Cnv2.Instruction.Task_ID;
                       "Transfer_To_ID_HMI(1)" := "Control_DB".LCnv_Sys[3].Cnv_Level[4].Cnv2.Instruction.Transfer_To_ID;
                       "Transfer_From_ID_HMI(1)" := "Control_DB".LCnv_Sys[3].Cnv_Level[4].Cnv2.Instruction.Transfer_From_ID;
                       "Pallet_Allignment_HMI(1)" := "Control_DB".LCnv_Sys[3].Cnv_Level[4].Cnv2.Instruction.Pallet_Allignment;
                   110503:
                       "Enable_HMI(1)" := "Control_DB".LCnv_Sys[3].Cnv_Level[5].Cnv2.Instruction.Enable;
                       "Mode_Change_HMI(1)" := "Control_DB".LCnv_Sys[3].Cnv_Level[5].Cnv2.Instruction.Mode_Change;
                       "Task_ID_HMI(1)" := "Control_DB".LCnv_Sys[3].Cnv_Level[5].Cnv2.Instruction.Task_ID;
                       "Transfer_To_ID_HMI(1)" := "Control_DB".LCnv_Sys[3].Cnv_Level[5].Cnv2.Instruction.Transfer_To_ID;
                       "Transfer_From_ID_HMI(1)" := "Control_DB".LCnv_Sys[3].Cnv_Level[5].Cnv2.Instruction.Transfer_From_ID;
                       "Pallet_Allignment_HMI(1)" := "Control_DB".LCnv_Sys[3].Cnv_Level[5].Cnv2.Instruction.Pallet_Allignment;
                   110603:
                       "Enable_HMI(1)" := "Control_DB".LCnv_Sys[3].Cnv_Level[6].Cnv2.Instruction.Enable;
                       "Mode_Change_HMI(1)" := "Control_DB".LCnv_Sys[3].Cnv_Level[6].Cnv2.Instruction.Mode_Change;
                       "Task_ID_HMI(1)" := "Control_DB".LCnv_Sys[3].Cnv_Level[6].Cnv2.Instruction.Task_ID;
                       "Transfer_To_ID_HMI(1)" := "Control_DB".LCnv_Sys[3].Cnv_Level[6].Cnv2.Instruction.Transfer_To_ID;
                       "Transfer_From_ID_HMI(1)" := "Control_DB".LCnv_Sys[3].Cnv_Level[6].Cnv2.Instruction.Transfer_From_ID;
                       "Pallet_Allignment_HMI(1)" := "Control_DB".LCnv_Sys[3].Cnv_Level[6].Cnv2.Instruction.Pallet_Allignment;
                   110703:
                       "Enable_HMI(1)" := "Control_DB".LCnv_Sys[3].Cnv_Level[7].Cnv2.Instruction.Enable;
                       "Mode_Change_HMI(1)" := "Control_DB".LCnv_Sys[3].Cnv_Level[7].Cnv2.Instruction.Mode_Change;
                       "Task_ID_HMI(1)" := "Control_DB".LCnv_Sys[3].Cnv_Level[7].Cnv2.Instruction.Task_ID;
                       "Transfer_To_ID_HMI(1)" := "Control_DB".LCnv_Sys[3].Cnv_Level[7].Cnv2.Instruction.Transfer_To_ID;
                       "Transfer_From_ID_HMI(1)" := "Control_DB".LCnv_Sys[3].Cnv_Level[7].Cnv2.Instruction.Transfer_From_ID;
                       "Pallet_Allignment_HMI(1)" := "Control_DB".LCnv_Sys[3].Cnv_Level[7].Cnv2.Instruction.Pallet_Allignment;
                   110803:
                       "Enable_HMI(1)" := "Control_DB".LCnv_Sys[3].Cnv_Level[8].Cnv2.Instruction.Enable;
                       "Mode_Change_HMI(1)" := "Control_DB".LCnv_Sys[3].Cnv_Level[8].Cnv2.Instruction.Mode_Change;
                       "Task_ID_HMI(1)" := "Control_DB".LCnv_Sys[3].Cnv_Level[8].Cnv2.Instruction.Task_ID;
                       "Transfer_To_ID_HMI(1)" := "Control_DB".LCnv_Sys[3].Cnv_Level[8].Cnv2.Instruction.Transfer_To_ID;
                       "Transfer_From_ID_HMI(1)" := "Control_DB".LCnv_Sys[3].Cnv_Level[8].Cnv2.Instruction.Transfer_From_ID;
                       "Pallet_Allignment_HMI(1)" := "Control_DB".LCnv_Sys[3].Cnv_Level[8].Cnv2.Instruction.Pallet_Allignment;
                       //CNV 2 - SYSTEM 4
                   110104:
                       "Enable_HMI(1)" := "Control_DB".LCnv_Sys[4].Cnv_Level[1].Cnv2.Instruction.Enable;
                       "Mode_Change_HMI(1)" := "Control_DB".LCnv_Sys[4].Cnv_Level[1].Cnv2.Instruction.Mode_Change;
                       "Task_ID_HMI(1)" := "Control_DB".LCnv_Sys[4].Cnv_Level[1].Cnv2.Instruction.Task_ID;
                       "Transfer_To_ID_HMI(1)" := "Control_DB".LCnv_Sys[4].Cnv_Level[1].Cnv2.Instruction.Transfer_To_ID;
                       "Transfer_From_ID_HMI(1)" := "Control_DB".LCnv_Sys[4].Cnv_Level[1].Cnv2.Instruction.Transfer_From_ID;
                       "Pallet_Allignment_HMI(1)" := "Control_DB".LCnv_Sys[4].Cnv_Level[1].Cnv2.Instruction.Pallet_Allignment;
                   110204:
                       "Enable_HMI(1)" := "Control_DB".LCnv_Sys[4].Cnv_Level[2].Cnv2.Instruction.Enable;
                       "Mode_Change_HMI(1)" := "Control_DB".LCnv_Sys[4].Cnv_Level[2].Cnv2.Instruction.Mode_Change;
                       "Task_ID_HMI(1)" := "Control_DB".LCnv_Sys[4].Cnv_Level[2].Cnv2.Instruction.Task_ID;
                       "Transfer_To_ID_HMI(1)" := "Control_DB".LCnv_Sys[4].Cnv_Level[2].Cnv2.Instruction.Transfer_To_ID;
                       "Transfer_From_ID_HMI(1)" := "Control_DB".LCnv_Sys[4].Cnv_Level[2].Cnv2.Instruction.Transfer_From_ID;
                       "Pallet_Allignment_HMI(1)" := "Control_DB".LCnv_Sys[4].Cnv_Level[2].Cnv2.Instruction.Pallet_Allignment;
                   110304:
                       "Enable_HMI(1)" := "Control_DB".LCnv_Sys[4].Cnv_Level[3].Cnv2.Instruction.Enable;
                       "Mode_Change_HMI(1)" := "Control_DB".LCnv_Sys[4].Cnv_Level[3].Cnv2.Instruction.Mode_Change;
                       "Task_ID_HMI(1)" := "Control_DB".LCnv_Sys[4].Cnv_Level[3].Cnv2.Instruction.Task_ID;
                       "Transfer_To_ID_HMI(1)" := "Control_DB".LCnv_Sys[4].Cnv_Level[3].Cnv2.Instruction.Transfer_To_ID;
                       "Transfer_From_ID_HMI(1)" := "Control_DB".LCnv_Sys[4].Cnv_Level[3].Cnv2.Instruction.Transfer_From_ID;
                       "Pallet_Allignment_HMI(1)" := "Control_DB".LCnv_Sys[4].Cnv_Level[3].Cnv2.Instruction.Pallet_Allignment;
                   110404:
                       "Enable_HMI(1)" := "Control_DB".LCnv_Sys[4].Cnv_Level[4].Cnv2.Instruction.Enable;
                       "Mode_Change_HMI(1)" := "Control_DB".LCnv_Sys[4].Cnv_Level[4].Cnv2.Instruction.Mode_Change;
                       "Task_ID_HMI(1)" := "Control_DB".LCnv_Sys[4].Cnv_Level[4].Cnv2.Instruction.Task_ID;
                       "Transfer_To_ID_HMI(1)" := "Control_DB".LCnv_Sys[4].Cnv_Level[4].Cnv2.Instruction.Transfer_To_ID;
                       "Transfer_From_ID_HMI(1)" := "Control_DB".LCnv_Sys[4].Cnv_Level[4].Cnv2.Instruction.Transfer_From_ID;
                       "Pallet_Allignment_HMI(1)" := "Control_DB".LCnv_Sys[4].Cnv_Level[4].Cnv2.Instruction.Pallet_Allignment;
                   110504:
                       "Enable_HMI(1)" := "Control_DB".LCnv_Sys[4].Cnv_Level[5].Cnv2.Instruction.Enable;
                       "Mode_Change_HMI(1)" := "Control_DB".LCnv_Sys[4].Cnv_Level[5].Cnv2.Instruction.Mode_Change;
                       "Task_ID_HMI(1)" := "Control_DB".LCnv_Sys[4].Cnv_Level[5].Cnv2.Instruction.Task_ID;
                       "Transfer_To_ID_HMI(1)" := "Control_DB".LCnv_Sys[4].Cnv_Level[5].Cnv2.Instruction.Transfer_To_ID;
                       "Transfer_From_ID_HMI(1)" := "Control_DB".LCnv_Sys[4].Cnv_Level[5].Cnv2.Instruction.Transfer_From_ID;
                       "Pallet_Allignment_HMI(1)" := "Control_DB".LCnv_Sys[4].Cnv_Level[5].Cnv2.Instruction.Pallet_Allignment;
                   110604:
                       "Enable_HMI(1)" := "Control_DB".LCnv_Sys[4].Cnv_Level[6].Cnv2.Instruction.Enable;
                       "Mode_Change_HMI(1)" := "Control_DB".LCnv_Sys[4].Cnv_Level[6].Cnv2.Instruction.Mode_Change;
                       "Task_ID_HMI(1)" := "Control_DB".LCnv_Sys[4].Cnv_Level[6].Cnv2.Instruction.Task_ID;
                       "Transfer_To_ID_HMI(1)" := "Control_DB".LCnv_Sys[4].Cnv_Level[6].Cnv2.Instruction.Transfer_To_ID;
                       "Transfer_From_ID_HMI(1)" := "Control_DB".LCnv_Sys[4].Cnv_Level[6].Cnv2.Instruction.Transfer_From_ID;
                       "Pallet_Allignment_HMI(1)" := "Control_DB".LCnv_Sys[4].Cnv_Level[6].Cnv2.Instruction.Pallet_Allignment;
                   110704:
                       "Enable_HMI(1)" := "Control_DB".LCnv_Sys[4].Cnv_Level[7].Cnv2.Instruction.Enable;
                       "Mode_Change_HMI(1)" := "Control_DB".LCnv_Sys[4].Cnv_Level[7].Cnv2.Instruction.Mode_Change;
                       "Task_ID_HMI(1)" := "Control_DB".LCnv_Sys[4].Cnv_Level[7].Cnv2.Instruction.Task_ID;
                       "Transfer_To_ID_HMI(1)" := "Control_DB".LCnv_Sys[4].Cnv_Level[7].Cnv2.Instruction.Transfer_To_ID;
                       "Transfer_From_ID_HMI(1)" := "Control_DB".LCnv_Sys[4].Cnv_Level[7].Cnv2.Instruction.Transfer_From_ID;
                       "Pallet_Allignment_HMI(1)" := "Control_DB".LCnv_Sys[4].Cnv_Level[7].Cnv2.Instruction.Pallet_Allignment;
                   110804:
                       "Enable_HMI(1)" := "Control_DB".LCnv_Sys[4].Cnv_Level[8].Cnv2.Instruction.Enable;
                       "Mode_Change_HMI(1)" := "Control_DB".LCnv_Sys[4].Cnv_Level[8].Cnv2.Instruction.Mode_Change;
                       "Task_ID_HMI(1)" := "Control_DB".LCnv_Sys[4].Cnv_Level[8].Cnv2.Instruction.Task_ID;
                       "Transfer_To_ID_HMI(1)" := "Control_DB".LCnv_Sys[4].Cnv_Level[8].Cnv2.Instruction.Transfer_To_ID;
                       "Transfer_From_ID_HMI(1)" := "Control_DB".LCnv_Sys[4].Cnv_Level[8].Cnv2.Instruction.Transfer_From_ID;
                       "Pallet_Allignment_HMI(1)" := "Control_DB".LCnv_Sys[4].Cnv_Level[8].Cnv2.Instruction.Pallet_Allignment;
                       //CNV 2 - SYSTEM 5
                   110105:
                       "Enable_HMI(1)" := "Control_DB".LCnv_Sys[5].Cnv_Level[1].Cnv2.Instruction.Enable;
                       "Mode_Change_HMI(1)" := "Control_DB".LCnv_Sys[5].Cnv_Level[1].Cnv2.Instruction.Mode_Change;
                       "Task_ID_HMI(1)" := "Control_DB".LCnv_Sys[5].Cnv_Level[1].Cnv2.Instruction.Task_ID;
                       "Transfer_To_ID_HMI(1)" := "Control_DB".LCnv_Sys[5].Cnv_Level[1].Cnv2.Instruction.Transfer_To_ID;
                       "Transfer_From_ID_HMI(1)" := "Control_DB".LCnv_Sys[5].Cnv_Level[1].Cnv2.Instruction.Transfer_From_ID;
                       "Pallet_Allignment_HMI(1)" := "Control_DB".LCnv_Sys[5].Cnv_Level[1].Cnv2.Instruction.Pallet_Allignment;
                   110205:
                       "Enable_HMI(1)" := "Control_DB".LCnv_Sys[5].Cnv_Level[2].Cnv2.Instruction.Enable;
                       "Mode_Change_HMI(1)" := "Control_DB".LCnv_Sys[5].Cnv_Level[2].Cnv2.Instruction.Mode_Change;
                       "Task_ID_HMI(1)" := "Control_DB".LCnv_Sys[5].Cnv_Level[2].Cnv2.Instruction.Task_ID;
                       "Transfer_To_ID_HMI(1)" := "Control_DB".LCnv_Sys[5].Cnv_Level[2].Cnv2.Instruction.Transfer_To_ID;
                       "Transfer_From_ID_HMI(1)" := "Control_DB".LCnv_Sys[5].Cnv_Level[2].Cnv2.Instruction.Transfer_From_ID;
                       "Pallet_Allignment_HMI(1)" := "Control_DB".LCnv_Sys[5].Cnv_Level[2].Cnv2.Instruction.Pallet_Allignment;
                   110305:
                       "Enable_HMI(1)" := "Control_DB".LCnv_Sys[5].Cnv_Level[3].Cnv2.Instruction.Enable;
                       "Mode_Change_HMI(1)" := "Control_DB".LCnv_Sys[5].Cnv_Level[3].Cnv2.Instruction.Mode_Change;
                       "Task_ID_HMI(1)" := "Control_DB".LCnv_Sys[5].Cnv_Level[3].Cnv2.Instruction.Task_ID;
                       "Transfer_To_ID_HMI(1)" := "Control_DB".LCnv_Sys[5].Cnv_Level[3].Cnv2.Instruction.Transfer_To_ID;
                       "Transfer_From_ID_HMI(1)" := "Control_DB".LCnv_Sys[5].Cnv_Level[3].Cnv2.Instruction.Transfer_From_ID;
                       "Pallet_Allignment_HMI(1)" := "Control_DB".LCnv_Sys[5].Cnv_Level[3].Cnv2.Instruction.Pallet_Allignment;
                   110405:
                       "Enable_HMI(1)" := "Control_DB".LCnv_Sys[5].Cnv_Level[4].Cnv2.Instruction.Enable;
                       "Mode_Change_HMI(1)" := "Control_DB".LCnv_Sys[5].Cnv_Level[4].Cnv2.Instruction.Mode_Change;
                       "Task_ID_HMI(1)" := "Control_DB".LCnv_Sys[5].Cnv_Level[4].Cnv2.Instruction.Task_ID;
                       "Transfer_To_ID_HMI(1)" := "Control_DB".LCnv_Sys[5].Cnv_Level[4].Cnv2.Instruction.Transfer_To_ID;
                       "Transfer_From_ID_HMI(1)" := "Control_DB".LCnv_Sys[5].Cnv_Level[4].Cnv2.Instruction.Transfer_From_ID;
                       "Pallet_Allignment_HMI(1)" := "Control_DB".LCnv_Sys[5].Cnv_Level[4].Cnv2.Instruction.Pallet_Allignment;
                   110505:
                       "Enable_HMI(1)" := "Control_DB".LCnv_Sys[5].Cnv_Level[5].Cnv2.Instruction.Enable;
                       "Mode_Change_HMI(1)" := "Control_DB".LCnv_Sys[5].Cnv_Level[5].Cnv2.Instruction.Mode_Change;
                       "Task_ID_HMI(1)" := "Control_DB".LCnv_Sys[5].Cnv_Level[5].Cnv2.Instruction.Task_ID;
                       "Transfer_To_ID_HMI(1)" := "Control_DB".LCnv_Sys[5].Cnv_Level[5].Cnv2.Instruction.Transfer_To_ID;
                       "Transfer_From_ID_HMI(1)" := "Control_DB".LCnv_Sys[5].Cnv_Level[5].Cnv2.Instruction.Transfer_From_ID;
                       "Pallet_Allignment_HMI(1)" := "Control_DB".LCnv_Sys[5].Cnv_Level[5].Cnv2.Instruction.Pallet_Allignment;
                   110605:
                       "Enable_HMI(1)" := "Control_DB".LCnv_Sys[5].Cnv_Level[6].Cnv2.Instruction.Enable;
                       "Mode_Change_HMI(1)" := "Control_DB".LCnv_Sys[5].Cnv_Level[6].Cnv2.Instruction.Mode_Change;
                       "Task_ID_HMI(1)" := "Control_DB".LCnv_Sys[5].Cnv_Level[6].Cnv2.Instruction.Task_ID;
                       "Transfer_To_ID_HMI(1)" := "Control_DB".LCnv_Sys[5].Cnv_Level[6].Cnv2.Instruction.Transfer_To_ID;
                       "Transfer_From_ID_HMI(1)" := "Control_DB".LCnv_Sys[5].Cnv_Level[6].Cnv2.Instruction.Transfer_From_ID;
                       "Pallet_Allignment_HMI(1)" := "Control_DB".LCnv_Sys[5].Cnv_Level[6].Cnv2.Instruction.Pallet_Allignment;
                   110705:
                       "Enable_HMI(1)" := "Control_DB".LCnv_Sys[5].Cnv_Level[7].Cnv2.Instruction.Enable;
                       "Mode_Change_HMI(1)" := "Control_DB".LCnv_Sys[5].Cnv_Level[7].Cnv2.Instruction.Mode_Change;
                       "Task_ID_HMI(1)" := "Control_DB".LCnv_Sys[5].Cnv_Level[7].Cnv2.Instruction.Task_ID;
                       "Transfer_To_ID_HMI(1)" := "Control_DB".LCnv_Sys[5].Cnv_Level[7].Cnv2.Instruction.Transfer_To_ID;
                       "Transfer_From_ID_HMI(1)" := "Control_DB".LCnv_Sys[5].Cnv_Level[7].Cnv2.Instruction.Transfer_From_ID;
                       "Pallet_Allignment_HMI(1)" := "Control_DB".LCnv_Sys[5].Cnv_Level[7].Cnv2.Instruction.Pallet_Allignment;
                   110805:
                       "Enable_HMI(1)" := "Control_DB".LCnv_Sys[5].Cnv_Level[8].Cnv2.Instruction.Enable;
                       "Mode_Change_HMI(1)" := "Control_DB".LCnv_Sys[5].Cnv_Level[8].Cnv2.Instruction.Mode_Change;
                       "Task_ID_HMI(1)" := "Control_DB".LCnv_Sys[5].Cnv_Level[8].Cnv2.Instruction.Task_ID;
                       "Transfer_To_ID_HMI(1)" := "Control_DB".LCnv_Sys[5].Cnv_Level[8].Cnv2.Instruction.Transfer_To_ID;
                       "Transfer_From_ID_HMI(1)" := "Control_DB".LCnv_Sys[5].Cnv_Level[8].Cnv2.Instruction.Transfer_From_ID;
                       "Pallet_Allignment_HMI(1)" := "Control_DB".LCnv_Sys[5].Cnv_Level[8].Cnv2.Instruction.Pallet_Allignment;
               END_CASE;
               "CNV_HMI".Charge_Commands[#HMI_No] := 0;
           END_IF;
       END_REGION

       REGION CHARGE DATA FROM HMI (AFTER CHARGE DATA)
           IF NOT "CNV_HMI".Charge_Commands[#HMI_No] AND NOT #R_Charge_Cnv_Commands.Q THEN
               CASE #"ID(1)" OF
                       //SYSTEM 1
                       //CNV 1
                   100101:
                       "Feed_BCNV_Cnv1(1)_1"(HMI_No := #HMI_No,
                                             System_No := #Sys_No,
                                             Level := 1,
                                             Light_Guard_IO:="LIGHT GUARDS C1101 - CH1",
                                             Light_Guard_Bypass=>"Light_Guard_Bypass(1)");
                   100201:
                       "Feed_BCNV_Cnv1(1)_1"(HMI_No := #HMI_No,
                                             System_No := #Sys_No,
                                             Level := 2,
                                             Light_Guard_IO:="LIGHT GUARDS C1101 - CH1",
                                             Light_Guard_Bypass=>"Light_Guard_Bypass(1)");
                   100301:
                       "Feed_BCNV_Cnv1(1)_1"(HMI_No := #HMI_No,
                                             System_No := #Sys_No,
                                             Level := 3,
                                             Light_Guard_IO:="LIGHT GUARDS C1101 - CH1",
                                             Light_Guard_Bypass=>"Light_Guard_Bypass(1)");
                   100401:
                       "Feed_BCNV_Cnv1(1)_1"(HMI_No := #HMI_No,
                                             System_No := #Sys_No,
                                             Level := 4,
                                             Light_Guard_IO:="LIGHT GUARDS C1101 - CH1",
                                             Light_Guard_Bypass=>"Light_Guard_Bypass(1)");
                   100501:
                       "Feed_BCNV_Cnv1(1)_1"(HMI_No := #HMI_No,
                                             System_No := #Sys_No,
                                             Level := 5,
                                             Light_Guard_IO:="LIGHT GUARDS C1101 - CH1",
                                             Light_Guard_Bypass=>"Light_Guard_Bypass(1)");
                   100601:
                       "Feed_BCNV_Cnv1(1)_1"(HMI_No := #HMI_No,
                                             System_No := #Sys_No,
                                             Level := 6,
                                             Light_Guard_IO:="LIGHT GUARDS C1101 - CH1",
                                             Light_Guard_Bypass=>"Light_Guard_Bypass(1)");
                   100701:
                       "Feed_BCNV_Cnv1(1)_1"(HMI_No := #HMI_No,
                                             System_No := #Sys_No,
                                             Level := 7,
                                             Light_Guard_IO:="LIGHT GUARDS C1101 - CH1",
                                             Light_Guard_Bypass=>"Light_Guard_Bypass(1)");
                   100801:
                       "Feed_BCNV_Cnv1(1)_1"(HMI_No := #HMI_No,
                                             System_No := #Sys_No,
                                             Level := 8,
                                             Light_Guard_IO:="LIGHT GUARDS C1101 - CH1",
                                             Light_Guard_Bypass=>"Light_Guard_Bypass(1)");
                       //CNV 2
                   110101:
                       "Feed_BCNV_Cnv2(1)_1"(HMI_No := #HMI_No,
                                             System_No := #Sys_No,
                                             Level := 1,
                                             Light_Guard_IO:="LIGHT GUARDS C1201 - CH1",
                                             Light_Guard_Bypass=>"Light_Guard_Bypass(1)");
                   110201:
                       "Feed_BCNV_Cnv2(1)_1"(HMI_No := #HMI_No,
                                             System_No := #Sys_No,
                                             Level := 2,
                                             Light_Guard_IO:="LIGHT GUARDS C1201 - CH1",
                                             Light_Guard_Bypass=>"Light_Guard_Bypass(1)");
                   110301:
                       "Feed_BCNV_Cnv2(1)_1"(HMI_No := #HMI_No,
                                             System_No := #Sys_No,
                                             Level := 3,
                                             Light_Guard_IO:="LIGHT GUARDS C1201 - CH1",
                                             Light_Guard_Bypass=>"Light_Guard_Bypass(1)");
                   110401:
                       "Feed_BCNV_Cnv2(1)_1"(HMI_No := #HMI_No,
                                             System_No := #Sys_No,
                                             Level := 4,
                                             Light_Guard_IO:="LIGHT GUARDS C1201 - CH1",
                                             Light_Guard_Bypass=>"Light_Guard_Bypass(1)");
                   110501:
                       "Feed_BCNV_Cnv2(1)_1"(HMI_No := #HMI_No,
                                             System_No := #Sys_No,
                                             Level := 5,
                                             Light_Guard_IO:="LIGHT GUARDS C1201 - CH1",
                                             Light_Guard_Bypass=>"Light_Guard_Bypass(1)");
                   110601:
                       "Feed_BCNV_Cnv2(1)_1"(HMI_No := #HMI_No,
                                             System_No := #Sys_No,
                                             Level := 6,
                                             Light_Guard_IO:="LIGHT GUARDS C1201 - CH1",
                                             Light_Guard_Bypass=>"Light_Guard_Bypass(1)");
                   110701:
                       "Feed_BCNV_Cnv2(1)_1"(HMI_No := #HMI_No,
                                             System_No := #Sys_No,
                                             Level := 7,
                                             Light_Guard_IO:="LIGHT GUARDS C1201 - CH1",
                                             Light_Guard_Bypass=>"Light_Guard_Bypass(1)");
                   110801:
                       "Feed_BCNV_Cnv2(1)_1"(HMI_No := #HMI_No,
                                             System_No := #Sys_No,
                                             Level := 8,
                                             Light_Guard_IO:="LIGHT GUARDS C1201 - CH1",
                                             Light_Guard_Bypass=>"Light_Guard_Bypass(1)");
                       //SYSTEM 2
                       //CNV 1
                   100102:
                       "Feed_BCNV_Cnv1(1)_1"(HMI_No := #HMI_No,
                                             System_No := 2,
                                             Level := 1,
                                             Light_Guard_IO:="LIGHT GUARDS C2101 - CH1",
                                             Light_Guard_Bypass=>"Light_Guard_Bypass(2)");
                   100202:
                       "Feed_BCNV_Cnv1(1)_1"(HMI_No := #HMI_No,
                                             System_No := 2,
                                             Level := 2,
                                             Light_Guard_IO:="LIGHT GUARDS C2101 - CH1",
                                             Light_Guard_Bypass=>"Light_Guard_Bypass(2)");
                   100302:
                       "Feed_BCNV_Cnv1(1)_1"(HMI_No := #HMI_No,
                                             System_No := 2,
                                             Level := 3,
                                             Light_Guard_IO:="LIGHT GUARDS C2101 - CH1",
                                             Light_Guard_Bypass=>"Light_Guard_Bypass(2)");
                   100402:
                       "Feed_BCNV_Cnv1(1)_1"(HMI_No := #HMI_No,
                                             System_No := 2,
                                             Level := 4,
                                             Light_Guard_IO:="LIGHT GUARDS C2101 - CH1",
                                             Light_Guard_Bypass=>"Light_Guard_Bypass(2)");
                   100502:
                       "Feed_BCNV_Cnv1(1)_1"(HMI_No := #HMI_No,
                                             System_No := 2,
                                             Level := 5,
                                             Light_Guard_IO:="LIGHT GUARDS C2101 - CH1",
                                             Light_Guard_Bypass=>"Light_Guard_Bypass(2)");
                   100602:
                       "Feed_BCNV_Cnv1(1)_1"(HMI_No := #HMI_No,
                                             System_No := 2,
                                             Level := 6,
                                             Light_Guard_IO:="LIGHT GUARDS C2101 - CH1",
                                             Light_Guard_Bypass=>"Light_Guard_Bypass(2)");
                   100702:
                       "Feed_BCNV_Cnv1(1)_1"(HMI_No := #HMI_No,
                                             System_No := 2,
                                             Level := 7,
                                             Light_Guard_IO:="LIGHT GUARDS C2101 - CH1",
                                             Light_Guard_Bypass=>"Light_Guard_Bypass(2)");
                   100802:
                       "Feed_BCNV_Cnv1(1)_1"(HMI_No := #HMI_No,
                                             System_No := 2,
                                             Level := 8,
                                             Light_Guard_IO:="LIGHT GUARDS C2101 - CH1",
                                             Light_Guard_Bypass=>"Light_Guard_Bypass(2)");
                       //CNV 2
                   110102:
                       "Feed_BCNV_Cnv2(1)_1"(HMI_No := #HMI_No,
                                             System_No := 2,
                                             Level := 1,
                                             Light_Guard_IO:="LIGHT GUARDS C2201 - CH1",
                                             Light_Guard_Bypass=>"Light_Guard_Bypass(2)");
                   110202:
                       "Feed_BCNV_Cnv2(1)_1"(HMI_No := #HMI_No,
                                             System_No := 2,
                                             Level := 2,
                                             Light_Guard_IO:="LIGHT GUARDS C2201 - CH1",
                                             Light_Guard_Bypass=>"Light_Guard_Bypass(2)");
                   110302:
                       "Feed_BCNV_Cnv2(1)_1"(HMI_No := #HMI_No,
                                             System_No := 2,
                                             Level := 3,
                                             Light_Guard_IO:="LIGHT GUARDS C2201 - CH1",
                                             Light_Guard_Bypass=>"Light_Guard_Bypass(2)");
                   110402:
                       "Feed_BCNV_Cnv2(1)_1"(HMI_No := #HMI_No,
                                             System_No := 2,
                                             Level := 4,
                                             Light_Guard_IO:="LIGHT GUARDS C2201 - CH1",
                                             Light_Guard_Bypass=>"Light_Guard_Bypass(2)");
                   110502:
                       "Feed_BCNV_Cnv2(1)_1"(HMI_No := #HMI_No,
                                             System_No := 2,
                                             Level := 5,
                                             Light_Guard_IO:="LIGHT GUARDS C2201 - CH1",
                                             Light_Guard_Bypass=>"Light_Guard_Bypass(2)");
                   110602:
                       "Feed_BCNV_Cnv2(1)_1"(HMI_No := #HMI_No,
                                             System_No := 2,
                                             Level := 6,
                                             Light_Guard_IO:="LIGHT GUARDS C2201 - CH1",
                                             Light_Guard_Bypass=>"Light_Guard_Bypass(2)");
                   110702:
                       "Feed_BCNV_Cnv2(1)_1"(HMI_No := #HMI_No,
                                             System_No := 2,
                                             Level := 7,
                                             Light_Guard_IO:="LIGHT GUARDS C2201 - CH1",
                                             Light_Guard_Bypass=>"Light_Guard_Bypass(2)");
                   110802:
                       "Feed_BCNV_Cnv2(1)_1"(HMI_No := #HMI_No,
                                             System_No := 2,
                                             Level := 8,
                                             Light_Guard_IO:="LIGHT GUARDS C2201 - CH1",
                                             Light_Guard_Bypass=>"Light_Guard_Bypass(2)");
                       //SYSTEM 3
                       //CNV 1
                   100103:
                       "Feed_BCNV_Cnv1(1)_1"(HMI_No := #HMI_No,
                                             System_No := 3,
                                             Level := 1,
                                             Light_Guard_IO:="LIGHT GUARDS C3101 - CH1",
                                             Light_Guard_Bypass=>"Light_Guard_Bypass(3)");
                   100203:
                       "Feed_BCNV_Cnv1(1)_1"(HMI_No := #HMI_No,
                                             System_No := 3,
                                             Level := 2,
                                             Light_Guard_IO:="LIGHT GUARDS C3101 - CH1",
                                             Light_Guard_Bypass=>"Light_Guard_Bypass(3)");
                   100303:
                       "Feed_BCNV_Cnv1(1)_1"(HMI_No := #HMI_No,
                                             System_No := 3,
                                             Level := 3,
                                             Light_Guard_IO:="LIGHT GUARDS C3101 - CH1",
                                             Light_Guard_Bypass=>"Light_Guard_Bypass(3)");
                   100403:
                       "Feed_BCNV_Cnv1(1)_1"(HMI_No := #HMI_No,
                                             System_No := 3,
                                             Level := 4,
                                             Light_Guard_IO:="LIGHT GUARDS C3101 - CH1",
                                             Light_Guard_Bypass=>"Light_Guard_Bypass(3)");
                   100503:
                       "Feed_BCNV_Cnv1(1)_1"(HMI_No := #HMI_No,
                                             System_No := 3,
                                             Level := 5,
                                             Light_Guard_IO:="LIGHT GUARDS C3101 - CH1",
                                             Light_Guard_Bypass=>"Light_Guard_Bypass(3)");
                   100603:
                       "Feed_BCNV_Cnv1(1)_1"(HMI_No := #HMI_No,
                                             System_No := 3,
                                             Level := 6,
                                             Light_Guard_IO:="LIGHT GUARDS C3101 - CH1",
                                             Light_Guard_Bypass=>"Light_Guard_Bypass(3)");
                   100703:
                       "Feed_BCNV_Cnv1(1)_1"(HMI_No := #HMI_No,
                                             System_No := 3,
                                             Level := 7,
                                             Light_Guard_IO:="LIGHT GUARDS C3101 - CH1",
                                             Light_Guard_Bypass=>"Light_Guard_Bypass(3)");
                   100803:
                       "Feed_BCNV_Cnv1(1)_1"(HMI_No := #HMI_No,
                                             System_No := 3,
                                             Level := 8,
                                             Light_Guard_IO:="LIGHT GUARDS C3101 - CH1",
                                             Light_Guard_Bypass=>"Light_Guard_Bypass(3)");
                       //CNV 2
                   110103:
                       "Feed_BCNV_Cnv2(1)_1"(HMI_No := #HMI_No,
                                             System_No := 3,
                                             Level := 1,
                                             Light_Guard_IO:="LIGHT GUARDS C3201 - CH1",
                                             Light_Guard_Bypass=>"Light_Guard_Bypass(3)");
                   110203:
                       "Feed_BCNV_Cnv2(1)_1"(HMI_No := #HMI_No,
                                             System_No := 3,
                                             Level := 2,
                                             Light_Guard_IO:="LIGHT GUARDS C3201 - CH1",
                                             Light_Guard_Bypass=>"Light_Guard_Bypass(3)");
                   110303:
                       "Feed_BCNV_Cnv2(1)_1"(HMI_No := #HMI_No,
                                             System_No := 3,
                                             Level := 3,
                                             Light_Guard_IO:="LIGHT GUARDS C3201 - CH1",
                                             Light_Guard_Bypass=>"Light_Guard_Bypass(3)");
                   110403:
                       "Feed_BCNV_Cnv2(1)_1"(HMI_No := #HMI_No,
                                             System_No := 3,
                                             Level := 4,
                                             Light_Guard_IO:="LIGHT GUARDS C3201 - CH1",
                                             Light_Guard_Bypass=>"Light_Guard_Bypass(3)");
                   110503:
                       "Feed_BCNV_Cnv2(1)_1"(HMI_No := #HMI_No,
                                             System_No := 3,
                                             Level := 5,
                                             Light_Guard_IO:="LIGHT GUARDS C3201 - CH1",
                                             Light_Guard_Bypass=>"Light_Guard_Bypass(3)");
                   110603:
                       "Feed_BCNV_Cnv2(1)_1"(HMI_No := #HMI_No,
                                             System_No := 3,
                                             Level := 6,
                                             Light_Guard_IO:="LIGHT GUARDS C3201 - CH1",
                                             Light_Guard_Bypass=>"Light_Guard_Bypass(3)");
                   110703:
                       "Feed_BCNV_Cnv2(1)_1"(HMI_No := #HMI_No,
                                             System_No := 3,
                                             Level := 7,
                                             Light_Guard_IO:="LIGHT GUARDS C3201 - CH1",
                                             Light_Guard_Bypass=>"Light_Guard_Bypass(3)");
                   110803:
                       "Feed_BCNV_Cnv2(1)_1"(HMI_No := #HMI_No,
                                             System_No := 3,
                                             Level := 8,
                                             Light_Guard_IO:="LIGHT GUARDS C3201 - CH1",
                                             Light_Guard_Bypass=>"Light_Guard_Bypass(3)");
                       //SYSTEM 4
                       //CNV 1
                   100104:
                       "Feed_BCNV_Cnv2(1)_1"(HMI_No := #HMI_No,
                                             System_No := 4,
                                             Level := 1,
                                             Light_Guard_IO:=TRUE,
                                             Light_Guard_Bypass=>#No_Light_Guard);
                   100204:
                       "Feed_BCNV_Cnv2(1)_1"(HMI_No := #HMI_No,
                                             System_No := 4,
                                             Level := 2,
                                             Light_Guard_IO:=TRUE,
                                             Light_Guard_Bypass=>#No_Light_Guard);
                   100304:
                       "Feed_BCNV_Cnv2(1)_1"(HMI_No := #HMI_No,
                                             System_No := 4,
                                             Level := 3,
                                             Light_Guard_IO:=TRUE,
                                             Light_Guard_Bypass=>#No_Light_Guard);
                   100404:
                       "Feed_BCNV_Cnv2(1)_1"(HMI_No := #HMI_No,
                                             System_No := 4,
                                             Level := 4,
                                             Light_Guard_IO:=TRUE,
                                             Light_Guard_Bypass=>#No_Light_Guard);
                   100504:
                       "Feed_BCNV_Cnv2(1)_1"(HMI_No := #HMI_No,
                                             System_No := 4,
                                             Level := 5,
                                             Light_Guard_IO:=TRUE,
                                             Light_Guard_Bypass=>#No_Light_Guard);
                   100604:
                       "Feed_BCNV_Cnv2(1)_1"(HMI_No := #HMI_No,
                                             System_No := 4,
                                             Level := 6,
                                             Light_Guard_IO:=TRUE,
                                             Light_Guard_Bypass=>#No_Light_Guard);
                   100704:
                       "Feed_BCNV_Cnv2(1)_1"(HMI_No := #HMI_No,
                                             System_No := 4,
                                             Level := 7,
                                             Light_Guard_IO:=TRUE,
                                             Light_Guard_Bypass=>#No_Light_Guard);
                   100804:
                       "Feed_BCNV_Cnv2(1)_1"(HMI_No := #HMI_No,
                                             System_No := 4,
                                             Level := 8,
                                             Light_Guard_IO:=TRUE,
                                             Light_Guard_Bypass=>#No_Light_Guard);
                       //SYSTEM 5
                       //CNV 1
                   100105:
                       "Feed_BCNV_Cnv2(1)_1"(HMI_No := #HMI_No,
                                             System_No := 5,
                                             Level := 1,
                                             Light_Guard_IO:=TRUE,
                                             Light_Guard_Bypass=>#No_Light_Guard);
                   100205:
                       "Feed_BCNV_Cnv2(1)_1"(HMI_No := #HMI_No,
                                             System_No := 5,
                                             Level := 2,
                                             Light_Guard_IO:=TRUE,
                                             Light_Guard_Bypass=>#No_Light_Guard);
                   100305:
                       "Feed_BCNV_Cnv2(1)_1"(HMI_No := #HMI_No,
                                             System_No := 5,
                                             Level := 3,
                                             Light_Guard_IO:=TRUE,
                                             Light_Guard_Bypass=>#No_Light_Guard);
                   100405:
                       "Feed_BCNV_Cnv2(1)_1"(HMI_No := #HMI_No,
                                             System_No := 5,
                                             Level := 4,
                                             Light_Guard_IO:=TRUE,
                                             Light_Guard_Bypass=>#No_Light_Guard);
                   100505:
                       "Feed_BCNV_Cnv2(1)_1"(HMI_No := #HMI_No,
                                             System_No := 5,
                                             Level := 5,
                                             Light_Guard_IO:=TRUE,
                                             Light_Guard_Bypass=>#No_Light_Guard);
                   100605:
                       "Feed_BCNV_Cnv2(1)_1"(HMI_No := #HMI_No,
                                             System_No := 5,
                                             Level := 6,
                                             Light_Guard_IO:=TRUE,
                                             Light_Guard_Bypass=>#No_Light_Guard);
                   100705:
                       "Feed_BCNV_Cnv2(1)_1"(HMI_No := #HMI_No,
                                             System_No := 5,
                                             Level := 7,
                                             Light_Guard_IO:=TRUE,
                                             Light_Guard_Bypass=>#No_Light_Guard);
                   100805:
                       "Feed_BCNV_Cnv2(1)_1"(HMI_No := #HMI_No,
                                             System_No := 5,
                                             Level := 8,
                                             Light_Guard_IO:=TRUE,
                                             Light_Guard_Bypass=>#No_Light_Guard);
               END_CASE;
           END_IF;
       END_REGION
   END_REGION


   //RESET CHARGE BITS
   #T_Reset_Charge.TON(IN := "VTD_HMI".Charge_VTD[#HMI_No] OR "CNV_HMI".Charge_Cnv[#HMI_No] OR "VTD_HMI".Charge_VTD_Commands[#HMI_No] OR "CNV_HMI".Charge_Commands[#HMI_No],
                       PT := T#2S);

   IF #T_Reset_Charge.Q THEN
       "VTD_HMI".Charge_VTD[#HMI_No] := FALSE;
       "CNV_HMI".Charge_Cnv[#HMI_No] := FALSE;
       "VTD_HMI".Charge_VTD_Commands[#HMI_No] := FALSE;
       "CNV_HMI".Charge_Commands[#HMI_No] := FALSE;
   END_IF;
END_FUNCTION_BLOCK

FUNCTION "FC_Orders" : Void   // FC96, SCL
{ S7_Optimized_Access := 'TRUE' }
VERSION : 0.1
// stored: AutoNumber true, IsIECCheckEnabled false, SetENOAutomatically false, UDAEnableTagReadback false
   VAR_INPUT
      Sys : UInt;
   END_VAR
   VAR_IN_OUT
      System : "System_UDT";
      Auto_Test : "Auto_Test";
      VTD_CurrentOrder : UDInt;
      Pallet_InOut_CurrentOrder : UDInt;
      Shuttle_InOut_CurrentOrder : UDInt;
      System_Busy : Bool;
   END_VAR
   VAR_TEMP
      i : Int;
      j : Int;
      EmptyOrder : "OrderTable_UDT";
   END_VAR
BEGIN
   IF "HMI_OrderTable".StartRow < 0 THEN
       "HMI_OrderTable".StartRow := 0;
   END_IF;
   IF "HMI_OrderTable".StartRow > 90 THEN
       "HMI_OrderTable".StartRow := 90;
   END_IF;

   //System - Order Table
   //Place Order manually
   IF "HMI_OrderTable".PlaceOrder_PB AND "HMI_OrderTable".PlacingNewOrder THEN
       "HMI_OrderTable".PlaceOrder_PB := FALSE;
       CASE "HMI_OrderTable".Device OF

           1:
               "HMI_OrderTable".OrderTable[0].Device := 'VTD';
           2:
               "HMI_OrderTable".OrderTable[0].Device := 'Pallet In Out';
           3:
               "HMI_OrderTable".OrderTable[0].Device := 'Shuttle In Out';
       END_CASE;
       IF "HMI_OrderTable".Device > 9 THEN
           "HMI_OrderTable".OrderTable[0].OPC_Control.Destination_Location := 0;
       END_IF;
       // "System_DB_VTD".OrderSent := "HMI_OrderTable".Device > 0;
       #System.StepTable[1] := "HMI_OrderTable".OrderTable[0];
       #System.StepTable[1].OrderNo := -1;
       #System.StepTable[1].StepNo := -1;
       #System.StepTable[1].PlaceTime := "Time".CurrentLocalTime;
       #System.StepTable[1].Status := 'Queued';
   END_IF;

   //Pause Order Push Button
   IF "HMI_OrderTable".PauseOrders_PB THEN
       "HMI_OrderTable".PauseOrders_PB := FALSE;
       #System.PauseOrders := TRUE;
   END_IF;
   //Resume Order Push Button
   IF "HMI_OrderTable".ResumeOrder_PB THEN
       "HMI_OrderTable".ResumeOrder_PB := FALSE;
       #System.ResumeOrders := TRUE;
   END_IF;
   //Cancel Order Push Button
   IF "HMI_OrderTable".CancelOrder_PB THEN
       "HMI_OrderTable".CancelOrder_PB := FALSE;
       #System.CancelOrders := TRUE;
   END_IF;

   //Cancel This Order Push Button
   IF "HMI_OrderTable".CancelThisOrder_PB THEN
       "HMI_OrderTable".CancelThisOrder_PB := FALSE;
       IF "HMI_OrderTable".OrderTable["HMI_OrderTable".PopUp_Index].Status = 'Error' THEN
           #System.OrderTable["HMI_OrderTable".PopUp_Index].Status := 'Error\Cancel';
           IF #System.CurrentOrder = "HMI_OrderTable".PopUp_Index THEN
               #System.CurrentOrder -= 1;
           END_IF;


           IF #System.OrderTable["HMI_OrderTable".PopUp_Index + "HMI_OrderTable".StartRow].Device = 'VTD' THEN
               #VTD_CurrentOrder := 0;
           ELSIF #System.OrderTable["HMI_OrderTable".PopUp_Index + "HMI_OrderTable".StartRow].Device = 'Pallet In Out' THEN
               #Pallet_InOut_CurrentOrder := 0;
           ELSIF #System.OrderTable["HMI_OrderTable".PopUp_Index + "HMI_OrderTable".StartRow].Device = 'Shuttle In Out' THEN
               #Shuttle_InOut_CurrentOrder := 0;
           END_IF;

       END_IF;

   END_IF;

   //Copy data
   FOR #i := 1 TO 9 DO
       #j := "HMI_OrderTable".StartRow + #i;
       "HMI_OrderTable".Index[#i] := #j;
       "HMI_OrderTable".OrderTable[#i] := #System.OrderTable[#j];
       //Color State
       IF "HMI_OrderTable".OrderTable[#i].Status = 'Queued' THEN
           "HMI_OrderTable".State[#i] := 1;
       ELSIF "HMI_OrderTable".OrderTable[#i].Status = 'Running' THEN
           "HMI_OrderTable".State[#i] := 2;
       ELSIF "HMI_OrderTable".OrderTable[#i].Status = 'Completed' THEN
           "HMI_OrderTable".State[#i] := 3;
       ELSIF "HMI_OrderTable".OrderTable[#i].Status = 'Error' THEN
           "HMI_OrderTable".State[#i] := 4;
       ELSIF "HMI_OrderTable".OrderTable[#i].Status = 'Paused' THEN
           "HMI_OrderTable".State[#i] := 5;
       ELSIF "HMI_OrderTable".OrderTable[#i].Status = 'Canceled' THEN
           "HMI_OrderTable".State[#i] := 6;
       ELSIF "HMI_OrderTable".OrderTable[#i].Status = 'Error\Cancel' THEN
           "HMI_OrderTable".State[#i] := 7;
       ELSE
           "HMI_OrderTable".State[#i] := 0;
       END_IF;
   END_FOR;

   IF NOT "HMI_OrderTable".PlacingNewOrder THEN
       "HMI_OrderTable".Device := 0;
   END_IF;

   //Error PopUp Window
   IF "HMI_OrderTable".PopUp_ErrorWindow_Active AND NOT "HMI_OrderTable".PlacingNewOrder THEN
       "HMI_OrderTable".OrderTable[0] := "HMI_OrderTable".OrderTable["HMI_OrderTable".PopUp_Index];
       IF "HMI_OrderTable".OrderTable[0].Status = 'Error' THEN
           "HMI_OrderTable".State[0] := 4;
       ELSIF "HMI_OrderTable".OrderTable[0].Status = 'Error\Cancel' THEN
           "HMI_OrderTable".State[0] := 7;
       ELSE
           "HMI_OrderTable".State[0] := 0;
       END_IF;
   ELSIF NOT "HMI_OrderTable".PopUp_ErrorWindow_Active AND NOT "HMI_OrderTable".PlacingNewOrder THEN
       "HMI_OrderTable".OrderTable[0] := #EmptyOrder;
   END_IF;

   REGION Testing area
       IF ("HMI_Box_Connected_1" = #System.Id OR ("HMI_Box_Connected_1" >= (#System.Id * 10) + 1 AND "HMI_Box_Connected_1" <= (#System.Id * 10) + 8)) OR
           ("HMI_Box_Connected_2" = #System.Id OR ("HMI_Box_Connected_1" >= (#System.Id * 10) + 1 AND "HMI_Box_Connected_1" <= (#System.Id * 10) + 8))
       THEN
           #System_Busy := TRUE;
       ELSE
           #System_Busy := FALSE;
           IF "Comissioning_Var" THEN
               //Visibilities
               //Running in auto mode
               IF #Auto_Test.Running AND NOT #Auto_Test.Manual AND NOT #Auto_Test.Pause THEN
                   "OrderTable_HMI"."Start Test Visibility" := FALSE;
                   "OrderTable_HMI"."Stop Test Visibility" := TRUE;
                   "OrderTable_HMI"."Pause Test Visibility" := TRUE;
                   "OrderTable_HMI"."Resume Visibility" := FALSE;
                   "OrderTable_HMI"."Clear Table Visibility" := FALSE;
                   "OrderTable_HMI"."Manual order Visibility" := FALSE;
                   //Running and paused
               ELSIF #Auto_Test.Running AND #Auto_Test.Pause AND NOT #Auto_Test.Manual THEN
                   "OrderTable_HMI"."Start Test Visibility" := FALSE;
                   "OrderTable_HMI"."Stop Test Visibility" := TRUE;
                   "OrderTable_HMI"."Pause Test Visibility" := FALSE;
                   "OrderTable_HMI"."Resume Visibility" := TRUE;
                   "OrderTable_HMI"."Clear Table Visibility" := FALSE;
                   "OrderTable_HMI"."Manual order Visibility" := FALSE;
                   //Running and Manual
               ELSIF #Auto_Test.Manual AND #Auto_Test.Running THEN
                   "OrderTable_HMI"."Start Test Visibility" := FALSE;
                   "OrderTable_HMI"."Stop Test Visibility" := FALSE;
                   "OrderTable_HMI"."Pause Test Visibility" := FALSE;
                   "OrderTable_HMI"."Resume Visibility" := FALSE;
                   "OrderTable_HMI"."Clear Table Visibility" := FALSE;
                   "OrderTable_HMI"."Manual order Visibility" := FALSE;
                   //Manual and not running
               ELSIF #Auto_Test.Manual AND NOT #Auto_Test.Running THEN
                   "OrderTable_HMI"."Start Test Visibility" := FALSE;
                   "OrderTable_HMI"."Stop Test Visibility" := FALSE;
                   "OrderTable_HMI"."Pause Test Visibility" := FALSE;
                   "OrderTable_HMI"."Resume Visibility" := FALSE;
                   "OrderTable_HMI"."Clear Table Visibility" := FALSE;
                   "OrderTable_HMI"."Manual order Visibility" := TRUE;
                   // not running, in automatic and no error
               ELSIF #Auto_Test.Automatic AND NOT #Auto_Test.Error AND #Auto_Test.State = 10 THEN
                   "OrderTable_HMI"."Start Test Visibility" := TRUE;
                   "OrderTable_HMI"."Stop Test Visibility" := FALSE;
                   "OrderTable_HMI"."Pause Test Visibility" := FALSE;
                   "OrderTable_HMI"."Resume Visibility" := FALSE;
                   "OrderTable_HMI"."Clear Table Visibility" := TRUE;
                   "OrderTable_HMI"."Manual order Visibility" := TRUE;
               ELSIF NOT #Auto_Test.Running THEN
                   "OrderTable_HMI"."Clear Table Visibility" := TRUE;
                   "OrderTable_HMI"."Manual order Visibility" := TRUE;
               END_IF;

               //PALLET TYPE VISIBILITY
               IF "OrderTable_HMI"."Pallet Type" = 1 THEN //CHEP
                   "OrderTable_HMI"."Tower 1 Visibility" := FALSE;
                   "OrderTable_HMI"."Tower 2 Visibility" := FALSE;
                   "OrderTable_HMI"."Extractor Visibility" := FALSE;
               ELSIF "OrderTable_HMI"."Pallet Type" = 2 THEN //EURO
                   "OrderTable_HMI"."Tower 1 Visibility" := TRUE;
                   "OrderTable_HMI"."Tower 2 Visibility" := TRUE;
                   "OrderTable_HMI"."Extractor Visibility" := TRUE;
               END_IF;

               IF #Auto_Test.Manual THEN
                   "OrderTable_HMI"."Tower Visibility" := TRUE;
                   "OrderTable_HMI"."Level Visibility" := TRUE;
                   "OrderTable_HMI"."ToExtractor Visibility" := TRUE;
                   "OrderTable_HMI".Auto_Settings_Visibility := FALSE;
                   IF #Auto_Test.Level <> 0 AND NOT #Auto_Test.Running THEN
                       "OrderTable_HMI"."Send VTD Order Visibility" := TRUE;
                   END_IF;
                   IF (("OrderTable_HMI"."Pallet Type" = 1) OR
                       ("OrderTable_HMI"."Pallet Type" = 2 AND "OrderTable_HMI".Tower = 1 AND "OrderTable_HMI"."Tower 1 Pallet Alignment" <> 0 AND "OrderTable_HMI".Transfer_From_To = 2) OR
                       ("OrderTable_HMI"."Pallet Type" = 2 AND "OrderTable_HMI".Tower = 2 AND "OrderTable_HMI"."Tower 1 Pallet Alignment" <> 0 AND "OrderTable_HMI".Transfer_From_To = 2) OR
                       ("OrderTable_HMI"."Pallet Type" = 2 AND "OrderTable_HMI"."Extractor Pallet Alignment" <> 0 AND "OrderTable_HMI".Transfer_From_To = 1))
                       AND
                       "OrderTable_HMI".Tower <> 0 AND "OrderTable_HMI".Transfer_From_To <> 0 AND NOT #Auto_Test.Running THEN
                       "OrderTable_HMI"."Send CNV Order Visibility" := TRUE;
                   ELSE
                       "OrderTable_HMI"."Send CNV Order Visibility" := FALSE;
                   END_IF;
               ELSE
                   "OrderTable_HMI"."Tower Visibility" := FALSE;
                   "OrderTable_HMI"."Level Visibility" := FALSE;
                   "OrderTable_HMI"."ToExtractor Visibility" := FALSE;
                   "OrderTable_HMI".Auto_Settings_Visibility := TRUE;
                   "OrderTable_HMI"."Send VTD Order Visibility" := FALSE;
                   "OrderTable_HMI"."Send CNV Order Visibility" := FALSE;
               END_IF;

               "OrderTable_HMI"."Pallet Type Visibility" := TRUE;
           ELSE
               "OrderTable_HMI"."Tower Visibility" := FALSE;
               "OrderTable_HMI"."Level Visibility" := FALSE;
               "OrderTable_HMI"."ToExtractor Visibility" := FALSE;
               "OrderTable_HMI".Auto_Settings_Visibility := FALSE;
               "OrderTable_HMI"."Send VTD Order Visibility" := FALSE;
               "OrderTable_HMI"."Send CNV Order Visibility" := FALSE;
               "OrderTable_HMI"."Pallet Type Visibility" := FALSE;
               "OrderTable_HMI"."Clear Table Visibility" := TRUE;
               "OrderTable_HMI"."Manual order Visibility" := FALSE;
           END_IF;

           //Buttons actions
           //START
           IF "OrderTable_HMI".Start THEN
               #Auto_Test.Start := TRUE;
           END_IF;

           //PAUSE
           IF "OrderTable_HMI".Pause THEN
               #Auto_Test.Pause := TRUE;
           END_IF;

           //STOP
           IF "OrderTable_HMI".Stop THEN
               #Auto_Test.Stop := TRUE;
           ELSE
               #Auto_Test.Stop := FALSE;
           END_IF;

           //RESUME
           IF "OrderTable_HMI".Resume THEN
               #Auto_Test.Pause := FALSE;
           END_IF;

           //MANUAL
           #Auto_Test.Manual := "OrderTable_HMI"."Manual order";

           //SEND VTD ORDER
           "R_Send_VTD_Order"(CLK := "OrderTable_HMI"."Send VTD Order");
           IF "R_Send_VTD_Order".Q THEN
               #Auto_Test.Send_VTD_Order := TRUE;
           END_IF;

           //SEND CNV ORDER
           "R_Send_CNV_Order"(CLK := "OrderTable_HMI"."Send CNV Order");
           IF "R_Send_CNV_Order".Q THEN
               #Auto_Test.Send_CNV_Order := TRUE;
           END_IF;

           //TEST SETTINGS
           //PALLET TYPE
           IF "OrderTable_HMI"."Pallet Type" = 1 THEN
               #Auto_Test."Pallet Type" := 'C';
           ELSIF "OrderTable_HMI"."Pallet Type" = 2 THEN
               #Auto_Test."Pallet Type" := 'E';
           ELSE
               #Auto_Test."Pallet Type" := ' ';
           END_IF;

           //PALLET ALIGNMENT TOWER 1
           IF "OrderTable_HMI"."Tower 1 Pallet Alignment" = 1 AND
               (("OrderTable_HMI".Transfer_From_To = 2 AND #Auto_Test.Manual) OR NOT #Auto_Test.Manual) THEN
               #Auto_Test."Tower 1 Pallet Alignment" := 'R';
               #Auto_Test.Pallet_Allignment := 'R';
           ELSIF "OrderTable_HMI"."Tower 1 Pallet Alignment" = 2 AND
               (("OrderTable_HMI".Transfer_From_To = 2 AND #Auto_Test.Manual) OR NOT #Auto_Test.Manual) THEN
               #Auto_Test."Tower 1 Pallet Alignment" := 'L';
               #Auto_Test.Pallet_Allignment := 'L';
           END_IF;

           //PALLET ALIGNMENT TOWER 2
           IF "OrderTable_HMI"."Tower 2 Pallet Alignment" = 1 AND
               (("OrderTable_HMI".Transfer_From_To = 2 AND #Auto_Test.Manual) OR NOT #Auto_Test.Manual) THEN
               #Auto_Test."Tower 2 Pallet Alignment" := 'R';
               #Auto_Test.Pallet_Allignment := 'R';
           ELSIF "OrderTable_HMI"."Tower 2 Pallet Alignment" = 2 AND
               (("OrderTable_HMI".Transfer_From_To = 2 AND #Auto_Test.Manual) OR NOT #Auto_Test.Manual) THEN
               #Auto_Test."Tower 2 Pallet Alignment" := 'L';
               #Auto_Test.Pallet_Allignment := 'L';
           END_IF;

           //PALLET ALIGNMENT ECONVEYOR
           IF "OrderTable_HMI"."Extractor Pallet Alignment" = 1 AND
               (("OrderTable_HMI".Transfer_From_To = 1 AND #Auto_Test.Manual) OR NOT #Auto_Test.Manual) THEN
               #Auto_Test."Extractor Pallet Alignment" := 'R';
               #Auto_Test.Pallet_Allignment := 'R';
           ELSIF "OrderTable_HMI"."Extractor Pallet Alignment" = 2 AND
               (("OrderTable_HMI".Transfer_From_To = 1 AND #Auto_Test.Manual) OR NOT #Auto_Test.Manual) THEN
               #Auto_Test."Extractor Pallet Alignment" := 'L';
               #Auto_Test.Pallet_Allignment := 'L';
           ELSIF "OrderTable_HMI"."Extractor Pallet Alignment" = 3 AND
               (("OrderTable_HMI".Transfer_From_To = 1 AND #Auto_Test.Manual) OR NOT #Auto_Test.Manual) THEN
               #Auto_Test."Extractor Pallet Alignment" := 'C';
               #Auto_Test.Pallet_Allignment := 'C';
           END_IF;

           //AUTOMATIC SETTING FOR BUTTON TRANSFER FROM_TO
           IF NOT "Control_DB".VTD_Sys[#Sys].Running AND "Control_DB".VTD_Sys[#Sys].Current_Level <> 0 THEN
               IF #Auto_Test.Tower = 1 AND "HMI_DB".ScreenNo_Main = 9 THEN
                   //CNV 1
                   IF "Control_DB".ECnv_Sys[#Sys].Cnv_Occupied AND NOT "Control_DB".LCnv_Sys[#Sys].Cnv_Level["Control_DB".VTD_Sys[#Sys].Current_Level].Cnv1.Cnv_Occupied AND
                       NOT "Control_DB".ECnv_Sys[#Sys].Running AND NOT "Control_DB".LCnv_Sys[#Sys].Cnv_Level["Control_DB".VTD_Sys[#Sys].Current_Level].Cnv1.Running THEN
                       #Auto_Test.Transfer_From_To := "OrderTable_HMI".Transfer_From_To := 2;//to buffer
                   ELSIF NOT "Control_DB".ECnv_Sys[#Sys].Cnv_Occupied AND "Control_DB".LCnv_Sys[#Sys].Cnv_Level["Control_DB".VTD_Sys[#Sys].Current_Level].Cnv1.Cnv_Occupied AND
                       NOT "Control_DB".ECnv_Sys[#Sys].Running AND NOT "Control_DB".LCnv_Sys[#Sys].Cnv_Level["Control_DB".VTD_Sys[#Sys].Current_Level].Cnv1.Running THEN
                       #Auto_Test.Transfer_From_To := "OrderTable_HMI".Transfer_From_To := 1;//to extractor
                   ELSE
                       #Auto_Test.Transfer_From_To := "OrderTable_HMI".Transfer_From_To;
                   END_IF;
                   //CNV 2
               ELSIF #Auto_Test.Tower = 2 AND "HMI_DB".ScreenNo_Main = 9 THEN   //CNV 2
                   IF "Control_DB".ECnv_Sys[#Sys].Cnv_Occupied AND NOT "Control_DB".LCnv_Sys[#Sys].Cnv_Level["Control_DB".VTD_Sys[#Sys].Current_Level].Cnv2.Cnv_Occupied AND
                       NOT "Control_DB".ECnv_Sys[#Sys].Running AND NOT "Control_DB".LCnv_Sys[#Sys].Cnv_Level["Control_DB".VTD_Sys[#Sys].Current_Level].Cnv2.Running THEN
                       #Auto_Test.Transfer_From_To := "OrderTable_HMI".Transfer_From_To := 2;
                   ELSIF NOT "Control_DB".ECnv_Sys[#Sys].Cnv_Occupied AND "Control_DB".LCnv_Sys[#Sys].Cnv_Level["Control_DB".VTD_Sys[#Sys].Current_Level].Cnv2.Cnv_Occupied AND
                       NOT "Control_DB".ECnv_Sys[#Sys].Running AND NOT "Control_DB".LCnv_Sys[#Sys].Cnv_Level["Control_DB".VTD_Sys[#Sys].Current_Level].Cnv2.Running THEN
                       #Auto_Test.Transfer_From_To := "OrderTable_HMI".Transfer_From_To := 1;
                   ELSE
                       #Auto_Test.Transfer_From_To := "OrderTable_HMI".Transfer_From_To;
                   END_IF;
               END_IF;
           END_IF;

           //LEVELS AND CYCLES
           #Auto_Test."From level" := "OrderTable_HMI"."From level";
           #Auto_Test."To level" := "OrderTable_HMI"."To level";
           #Auto_Test."Testing Time" := "OrderTable_HMI"."Testing Time";
           #Auto_Test."Numer of cycles" := "OrderTable_HMI"."Numer of cycles";
           #Auto_Test.Level := "OrderTable_HMI".Level;
           #Auto_Test.Tower := "OrderTable_HMI".Tower;
           "OrderTable_HMI"."Time Running" := DINT_TO_UINT(TIME_TO_DINT(#Auto_Test.Time_Runnng) / 60000);
           "OrderTable_HMI".Actual_Cycle := UINT_TO_BYTE(#Auto_Test.N_Cycles);
       END_IF;
   END_REGION ;
END_FUNCTION

FUNCTION "FC_Orders_1" : Void   // FC97, SCL
{ S7_Optimized_Access := 'TRUE' }
VERSION : 0.1
// stored: AutoNumber true, IsIECCheckEnabled false, SetENOAutomatically false, UDAEnableTagReadback false
   VAR_INPUT
      Sys : UInt;
   END_VAR
   VAR_IN_OUT
      System : "System_UDT";
      VTD_CurrentOrder : UDInt;
      Pallet_InOut_CurrentOrder : UDInt;
      Shuttle_InOut_CurrentOrder : UDInt;
   END_VAR
   VAR_TEMP
      i : Int;
      j : Int;
      EmptyOrder : "OrderTable_UDT";
   END_VAR
BEGIN
   IF "HMI_OrderTable_1".StartRow < 0 THEN
       "HMI_OrderTable_1".StartRow := 0;
   END_IF;
   IF "HMI_OrderTable_1".StartRow > 90 THEN
       "HMI_OrderTable_1".StartRow := 90;
   END_IF;

   //System - Order Table
   //Place Order manually
   IF "HMI_OrderTable_1".PlaceOrder_PB AND "HMI_OrderTable_1".PlacingNewOrder THEN
       "HMI_OrderTable_1".PlaceOrder_PB := FALSE;
       CASE "HMI_OrderTable_1".Device OF

           1:
               "HMI_OrderTable_1".OrderTable[0].Device := 'VTD';
           2:
               "HMI_OrderTable_1".OrderTable[0].Device := 'Pallet In Out';
           3:
               "HMI_OrderTable_1".OrderTable[0].Device := 'Shuttle In Out';
       END_CASE;
       IF "HMI_OrderTable_1".Device > 9 THEN
           "HMI_OrderTable_1".OrderTable[0].OPC_Control.Destination_Location := 0;
       END_IF;
       // "System_DB_VTD".OrderSent := "HMI_OrderTable_1".Device > 0;
       #System.StepTable[1] := "HMI_OrderTable_1".OrderTable[0];
       #System.StepTable[1].OrderNo := -1;
       #System.StepTable[1].StepNo := -1;
       #System.StepTable[1].PlaceTime := "Time".CurrentLocalTime;
       #System.StepTable[1].Status := 'Queued';
   END_IF;

   //Pause Order Push Button
   IF "HMI_OrderTable_1".PauseOrders_PB THEN
       "HMI_OrderTable_1".PauseOrders_PB := FALSE;
       #System.PauseOrders := TRUE;
   END_IF;
   //Resume Order Push Button
   IF "HMI_OrderTable_1".ResumeOrder_PB THEN
       "HMI_OrderTable_1".ResumeOrder_PB := FALSE;
       #System.ResumeOrders := TRUE;
   END_IF;
   //Cancel Order Push Button
   IF "HMI_OrderTable_1".CancelOrder_PB THEN
       "HMI_OrderTable_1".CancelOrder_PB := FALSE;
       #System.CancelOrders := TRUE;
   END_IF;

   //Cancel This Order Push Button
   IF "HMI_OrderTable_1".CancelThisOrder_PB THEN
       "HMI_OrderTable_1".CancelThisOrder_PB := FALSE;
       IF "HMI_OrderTable_1".OrderTable["HMI_OrderTable_1".PopUp_Index].Status = 'Error' THEN
           #System.OrderTable["HMI_OrderTable_1".PopUp_Index].Status := 'Error\Cancel';
           IF #System.CurrentOrder = "HMI_OrderTable_1".PopUp_Index THEN
               #System.CurrentOrder -= 1;
           END_IF;


           IF #System.OrderTable["HMI_OrderTable_1".PopUp_Index + "HMI_OrderTable_1".StartRow].Device = 'VTD' THEN
               #VTD_CurrentOrder := 0;
           ELSIF #System.OrderTable["HMI_OrderTable_1".PopUp_Index + "HMI_OrderTable_1".StartRow].Device = 'Pallet In Out' THEN
               #Pallet_InOut_CurrentOrder := 0;
           ELSIF #System.OrderTable["HMI_OrderTable_1".PopUp_Index + "HMI_OrderTable_1".StartRow].Device = 'Shuttle In Out' THEN
               #Shuttle_InOut_CurrentOrder := 0;
           END_IF;

       END_IF;

   END_IF;

   //Copy data
   FOR #i := 1 TO 9 DO
       #j := "HMI_OrderTable_1".StartRow + #i;
       "HMI_OrderTable_1".Index[#i] := #j;
       "HMI_OrderTable_1".OrderTable[#i] := #System.OrderTable[#j];
       //Color State
       IF "HMI_OrderTable_1".OrderTable[#i].Status = 'Queued' THEN
           "HMI_OrderTable_1".State[#i] := 1;
       ELSIF "HMI_OrderTable_1".OrderTable[#i].Status = 'Running' THEN
           "HMI_OrderTable_1".State[#i] := 2;
       ELSIF "HMI_OrderTable_1".OrderTable[#i].Status = 'Completed' THEN
           "HMI_OrderTable_1".State[#i] := 3;
       ELSIF "HMI_OrderTable_1".OrderTable[#i].Status = 'Error' THEN
           "HMI_OrderTable_1".State[#i] := 4;
       ELSIF "HMI_OrderTable_1".OrderTable[#i].Status = 'Paused' THEN
           "HMI_OrderTable_1".State[#i] := 5;
       ELSIF "HMI_OrderTable_1".OrderTable[#i].Status = 'Canceled' THEN
           "HMI_OrderTable_1".State[#i] := 6;
       ELSIF "HMI_OrderTable_1".OrderTable[#i].Status = 'Error\Cancel' THEN
           "HMI_OrderTable_1".State[#i] := 7;
       ELSE
           "HMI_OrderTable_1".State[#i] := 0;
       END_IF;
   END_FOR;

   IF NOT "HMI_OrderTable_1".PlacingNewOrder THEN
       "HMI_OrderTable_1".Device := 0;
   END_IF;

   //Error PopUp Window
   IF "HMI_OrderTable_1".PopUp_ErrorWindow_Active AND NOT "HMI_OrderTable_1".PlacingNewOrder THEN
       "HMI_OrderTable_1".OrderTable[0] := "HMI_OrderTable_1".OrderTable["HMI_OrderTable_1".PopUp_Index];
       IF "HMI_OrderTable_1".OrderTable[0].Status = 'Error' THEN
           "HMI_OrderTable_1".State[0] := 4;
       ELSIF "HMI_OrderTable_1".OrderTable[0].Status = 'Error\Cancel' THEN
           "HMI_OrderTable_1".State[0] := 7;
       ELSE
           "HMI_OrderTable_1".State[0] := 0;
       END_IF;
   ELSIF NOT "HMI_OrderTable_1".PopUp_ErrorWindow_Active AND NOT "HMI_OrderTable_1".PlacingNewOrder THEN
       "HMI_OrderTable_1".OrderTable[0] := #EmptyOrder;
   END_IF;
END_FUNCTION

FUNCTION "FC_Orders_2" : Void   // FC98, SCL
{ S7_Optimized_Access := 'TRUE' }
VERSION : 0.1
// stored: AutoNumber true, IsIECCheckEnabled false, SetENOAutomatically false, UDAEnableTagReadback false
   VAR_INPUT
      Sys : UInt;
   END_VAR
   VAR_IN_OUT
      System : "System_UDT";
      Auto_Test : "Auto_Test_1";
      VTD_CurrentOrder : UDInt;
      Pallet_InOut_CurrentOrder : UDInt;
      Shuttle_InOut_CurrentOrder : UDInt;
      System_Busy : Bool;
   END_VAR
   VAR_TEMP
      i : Int;
      j : Int;
      EmptyOrder : "OrderTable_UDT";
   END_VAR
BEGIN
   IF "HMI_OrderTable".StartRow < 0 THEN
       "HMI_OrderTable".StartRow := 0;
   END_IF;
   IF "HMI_OrderTable".StartRow > 90 THEN
       "HMI_OrderTable".StartRow := 90;
   END_IF;

   //System - Order Table
   //Place Order manually
   IF "HMI_OrderTable".PlaceOrder_PB AND "HMI_OrderTable".PlacingNewOrder THEN
       "HMI_OrderTable".PlaceOrder_PB := FALSE;
       CASE "HMI_OrderTable".Device OF

           1:
               "HMI_OrderTable".OrderTable[0].Device := 'VTD';
           2:
               "HMI_OrderTable".OrderTable[0].Device := 'Pallet In Out';
           3:
               "HMI_OrderTable".OrderTable[0].Device := 'Shuttle In Out';
       END_CASE;
       IF "HMI_OrderTable".Device > 9 THEN
           "HMI_OrderTable".OrderTable[0].OPC_Control.Destination_Location := 0;
       END_IF;
       // "System_DB_VTD".OrderSent := "HMI_OrderTable".Device > 0;
       #System.StepTable[1] := "HMI_OrderTable".OrderTable[0];
       #System.StepTable[1].OrderNo := -1;
       #System.StepTable[1].StepNo := -1;
       #System.StepTable[1].PlaceTime := "Time".CurrentLocalTime;
       #System.StepTable[1].Status := 'Queued';
   END_IF;

   //Pause Order Push Button
   IF "HMI_OrderTable".PauseOrders_PB THEN
       "HMI_OrderTable".PauseOrders_PB := FALSE;
       #System.PauseOrders := TRUE;
   END_IF;
   //Resume Order Push Button
   IF "HMI_OrderTable".ResumeOrder_PB THEN
       "HMI_OrderTable".ResumeOrder_PB := FALSE;
       #System.ResumeOrders := TRUE;
   END_IF;
   //Cancel Order Push Button
   IF "HMI_OrderTable".CancelOrder_PB THEN
       "HMI_OrderTable".CancelOrder_PB := FALSE;
       #System.CancelOrders := TRUE;
   END_IF;

   //Cancel This Order Push Button
   IF "HMI_OrderTable".CancelThisOrder_PB THEN
       "HMI_OrderTable".CancelThisOrder_PB := FALSE;
       IF "HMI_OrderTable".OrderTable["HMI_OrderTable".PopUp_Index].Status = 'Error' THEN
           #System.OrderTable["HMI_OrderTable".PopUp_Index].Status := 'Error\Cancel';
           IF #System.CurrentOrder = "HMI_OrderTable".PopUp_Index THEN
               #System.CurrentOrder -= 1;
           END_IF;


           IF #System.OrderTable["HMI_OrderTable".PopUp_Index + "HMI_OrderTable".StartRow].Device = 'VTD' THEN
               #VTD_CurrentOrder := 0;
           ELSIF #System.OrderTable["HMI_OrderTable".PopUp_Index + "HMI_OrderTable".StartRow].Device = 'Pallet In Out' THEN
               #Pallet_InOut_CurrentOrder := 0;
           ELSIF #System.OrderTable["HMI_OrderTable".PopUp_Index + "HMI_OrderTable".StartRow].Device = 'Shuttle In Out' THEN
               #Shuttle_InOut_CurrentOrder := 0;
           END_IF;

       END_IF;

   END_IF;

